IF FStep = CompleteState THEN
    FCompletedSequence := FCaptureStatus.SequenceId;
END_IF;
IF FStep >= LateChildProgress THEN
    FStatusRefreshMatches := (Snapshot.Execution.State = E_State.Completed)
        AND Snapshot.Execution.Completed AND NOT Snapshot.Execution.Ready
        AND (Snapshot.Execution.Result = FExpectedFinalResult)
        AND (Snapshot.TestCaseCountTotal = 2) AND (Snapshot.TestCaseCountRunning = 0);
    IF LateResetChildren THEN
        FStatusRefreshMatches := FStatusRefreshMatches AND Snapshot.Execution.Error
            AND (Snapshot.TestCaseCountCompleted = 1) AND (Snapshot.TestCaseCountError = 1)
            AND (Snapshot.TestCaseCountIdle = 1) AND (Snapshot.TestCaseCountPassed = 0);
    ELSE
        FStatusRefreshMatches := FStatusRefreshMatches AND NOT Snapshot.Execution.Error
            AND (Snapshot.TestCaseCountCompleted = 2) AND (Snapshot.TestCaseCountPassed = 2)
            AND (Snapshot.TestCaseCountIdle = 0) AND (Snapshot.TestCaseCountError = 0);
    END_IF;
    FPublicationMatches := FPublicationMatches AND (FCaptureStatus.SequenceId = FCompletedSequence);
END_IF;
IF (FStep = ReleaseReservations) OR (FStep = QuietAfterRelease)
    OR ((FStep = ResetOutcome) AND NOT LateResetChildren) THEN
    Released := FSubject.FreeReservedEvents();
    FCleanupMatches := Released
        AND (FSubject.ReservedEntryCount = 0) AND (FCapture.ReservedEntryCount = 0)
        AND (FSubject.State = ExpectedState) AND (FSubject.Result = ExpectedResult);
END_IF;

IF FExpectCompletion THEN
    FPublicationMatches := FPublicationMatches AND (FCaptureStatus.SequenceId = FCompletedSequence);
END_IF;
END_METHOD

END_FUNCTION_BLOCK

// ---- SelfTests/TestCases/TestSuite_TestSuiteLifecycle/Test_SuiteReservationRelease.TcPOU
{region 'Documentation'}
(*!
<summary>Verifies Suite release delegation, partial success, zero-own-budget cleanup and idempotent retry.</summary>
<description>

Boundary under test

The Suite uses the real local EventBuffer for its own contribution. Controlled children retain
local reservation markers only; they deliberately do not reproduce global reservation accounting.
The test checks that every child is called even if the first rejects release and that the Suite
still releases its own contribution. Global child-budget arithmetic belongs to capacity tests.

Retry and lifecycle

A failed child keeps its marker. A later successful retry releases it without re-releasing
already cleared contributions. Cleanup also visits children when the Suite's own count is zero.
None of these calls may issue child lifecycle requests, change owner state or restart execution.
</description>
*)
{endregion}
FUNCTION_BLOCK Test_SuiteReservationRelease EXTENDS TestCaseBase
VAR
    FSubjectParent : I_RunControl;
    FSubject : TestSuiteLifecycleProbe;
    FHelper : SuiteOrchestratorDouble;
    FCapture : EventBuffer;
    FEvents : ARRAY[1..CaptureLength] OF ST_Event;
    FCaptureFifo : ST_FifoStatus;
    FCaptureStatus : ST_EventBufferStatus;
    FChildView : ST_OrchestrationObservation;
    FStep : INT;
    FStepChecked : BOOL;
    FQuietSequence : UDINT;
    FDelegation : AssertTrue;
    FDelegationMatches : BOOL := TRUE;
    FOwnRelease : AssertTrue;
    FOwnReleaseMatches : BOOL := TRUE;
    FIdempotence : AssertTrue;
    FIdempotenceMatches : BOOL := TRUE;
    FNoLifecycleEffects : AssertTrue;
    FNoLifecycleEffectsMatches : BOOL := TRUE;
    FChildCalls : AssertTrue;
    FChildCallsMatches : BOOL := TRUE;
END_VAR
VAR CONSTANT
    CaptureLength : UINT := 64;
    ReservationMarker : UINT := 1;
    Setup : INT := 0;
    ResetRequested : INT := 1;
    FinishReset : INT := 2;
    ReserveAll : INT := 3;
    PartialRelease : INT := 4;
    RetryRelease : INT := 5;
    ReleaseWithZeroOwnCount : INT := 6;
    RepeatRelease : INT := 7;
    Done : INT := 8;
END_VAR

SUPER^();

{region 'Documentation'}
(*!
<summary>Contributes only the checking Assertions, not the intentionally controlled subject results.</summary>
*)
{endregion}
METHOD PROTECTED AggregateResults
VAR_INPUT
    Aggregator : I_ResultAggregator; //! Borrowed result sink owned by the outer Test Case; add this test's checking Assertions without resetting or retaining the sink.
END_VAR
Aggregator.AddProvider(Provider := FDelegation);
Aggregator.AddProvider(Provider := FOwnRelease);
Aggregator.AddProvider(Provider := FIdempotence);
Aggregator.AddProvider(Provider := FNoLifecycleEffects);
Aggregator.AddProvider(Provider := FChildCalls);
END_METHOD

{region 'Documentation'}
(*!
<summary>Supplies only the root identity; the root never executes this isolated subject.</summary>
*)
{endregion}
METHOD PUBLIC BindSubjectParent
VAR_INPUT
    Parent : I_RunControl; //! Borrowed identity parent retained for isolated subject initialization; keep the Run-Control alive through subject use.
END_VAR
FSubjectParent := Parent;
END_METHOD

{region 'Documentation'}
(*!
<summary>Initializes the checking Assertions; the scenario explicitly initializes its isolated subject.</summary>
*)
{endregion}
METHOD PROTECTED Configure
FPreparationStateCount := 0;
FTestStateCount := 1;
FDelegation.Initialize(Parent := THIS^,
    AssertionName := 'Delegation');
FOwnRelease.Initialize(Parent := THIS^,
    AssertionName := 'OwnRelease');
FIdempotence.Initialize(Parent := THIS^,
    AssertionName := 'Idempotence');
FNoLifecycleEffects.Initialize(Parent := THIS^,
    AssertionName := 'NoLifecycleEffects');
FChildCalls.Initialize(Parent := THIS^,
    AssertionName := 'ChildCalls');
END_METHOD

{region 'Documentation'}
(*!
<summary>No asynchronous test resource remains to stop.</summary>
*)
{endregion}
METHOD PROTECTED ProcessAbort
VAR_INPUT
    Enable : BOOL; //! Phase permission supplied by the owning Test Case; FALSE does not authorize progression, while observation may continue.
END_VAR
IF Enable THEN
    CompleteAbort();
END_IF;
END_METHOD

{region 'Documentation'}
(*!
<summary>Checks each cleanup checkpoint before advancing; failures remain latched.</summary>
*)
{endregion}
METHOD PROTECTED ProcessAssertions
VAR_INPUT
    Enable : BOOL; //! Phase permission supplied by the owning Test Case; FALSE does not authorize progression, while observation may continue.
END_VAR
FDelegation(Enable := Enable,
    State := State,
    IN := FDelegationMatches);
FOwnRelease(Enable := Enable,
    State := State,
    IN := FOwnReleaseMatches);
FIdempotence(Enable := Enable,
    State := State,
    IN := FIdempotenceMatches);
FNoLifecycleEffects(Enable := Enable,
    State := State,
    IN := FNoLifecycleEffectsMatches);
FChildCalls(Enable := Enable,
    State := State,
    IN := FChildCallsMatches);
IF Enable THEN
    FStepChecked := TRUE;
END_IF;
END_METHOD

{region 'Documentation'}
(*!
<summary>No resource Preparation is required for this controlled owner scenario.</summary>
*)
{endregion}
METHOD PROTECTED ProcessPreparations
VAR_INPUT
    // SA0033: Required override; the scenario has no Preparation phase.
    {attribute 'analysis' := '-33'}
    Enable : BOOL; //! Phase permission supplied by the owning Test Case; FALSE does not authorize progression, while observation may continue.
END_VAR
END_METHOD

{region 'Documentation'}
(*!
<summary>Restarts the test script and clears checking Assertions; subject setup belongs to the next test attempt.</summary>
*)
{endregion}
METHOD PROTECTED ProcessReset
FStep := Setup;
FStepChecked := FALSE;
FQuietSequence := 0;
FDelegationMatches := TRUE;
FOwnReleaseMatches := TRUE;
FIdempotenceMatches := TRUE;
FNoLifecycleEffectsMatches := TRUE;
FChildCallsMatches := TRUE;
FDelegation.Reset();
FOwnRelease.Reset();
FIdempotence.Reset();
FNoLifecycleEffects.Reset();
FChildCalls.Reset();
CompleteReset();
END_METHOD

{region 'Documentation'}
(*!
<summary>Advances the explicit test script with at most one subject FB call per active PLC cycle.</summary>
*)
{endregion}
METHOD PROTECTED ProcessTests
VAR_INPUT
    Enable : BOOL; //! Phase permission supplied by the owning Test Case; FALSE does not authorize progression, while observation may continue.
END_VAR
IF NOT Enable THEN
    RETURN;
END_IF;
IF FStepChecked THEN
    FStep := FStep + 1;
    FStepChecked := FALSE;
END_IF;
IF FStep = Done THEN
    CompleteTests();
    RETURN;
END_IF;
RunStep();
END_METHOD

{region 'Documentation'}
(*!
<summary>Exercises a bounded cleanup sequence in Idle, recording each concrete child release attempt.</summary>
*)
{endregion}
METHOD PRIVATE RunStep
VAR
    Config : ST_TestSuiteConfig;
    FirstChild : I_TestCase;
    SecondChild : I_TestCase;
    FirstCalls : ST_OrchestrationCalls;
    SecondCalls : ST_OrchestrationCalls;
    ExpectedState : E_State;
    ExpectedTask : E_OrchestratorTask;
    Released : BOOL;
END_VAR
IF FStep = Setup THEN
    IF NOT FCapture.Initialize(Buffer := FEvents,
        FifoControl := FCaptureFifo,
        Status := FCaptureStatus) THEN
        Error(Message := 'Suite release capture could not be initialized.');
        RETURN;
    END_IF;
    FHelper.BeginScenario();
    FSubject.Bind(Publisher := FCapture,
        Helper := FHelper);
    IF NOT FSubject.Initialize(Parent := FSubjectParent,
        SuiteName := 'ReleaseSubject',
        Config := Config) THEN
        Error(Message := 'Suite release subject could not be initialized.');
        RETURN;
    END_IF;
END_IF;
FirstChild := FSubject.GetTestCase(Index := FSubject.ChildArrayLowerBound);
SecondChild := FSubject.GetTestCase(Index := FSubject.ChildArrayLowerBound + 1);
ExpectedState := E_State.Idle;
ExpectedTask := E_OrchestratorTask.Idle;

CASE FStep OF
    Setup:
        FChildView.State := E_State.Uninitialized;
        FChildView.Result := E_Result.NotEvaluated;
        FChildView.Ready := FALSE;
        FChildView.Complete := FALSE;
        ExpectedState := E_State.Uninitialized;

    ResetRequested:
        IF FSubject.ReserveResetEvents() <> E_EventReservationResult.Accepted THEN
            Error(Message := 'Suite release fixture Reset reservation was rejected.');
            RETURN;
        END_IF;
        FSubject.RequestReset();
        FChildView.State := E_State.Reset;
        ExpectedState := E_State.Reset;
        ExpectedTask := E_OrchestratorTask.Reset;

    FinishReset:
        FHelper.SetObservation(Ready := TRUE,
            ResetFinished := TRUE);
        FChildView.State := E_State.Idle;
        FChildView.Ready := TRUE;

    ReserveAll:
        IF FSubject.ReserveExecutionEvents() <> E_EventReservationResult.Accepted THEN
            Error(Message := 'Suite release fixture execution reservation was rejected.');
            RETURN;
        END_IF;
        IF FirstChild.ReserveExecutionEvents() <> E_EventReservationResult.Accepted THEN
            Error(Message := 'First controlled child reservation was rejected.');
            RETURN;
        END_IF;
        IF SecondChild.ReserveExecutionEvents() <> E_EventReservationResult.Accepted THEN
            Error(Message := 'Second controlled child reservation was rejected.');
            RETURN;
        END_IF;
        FOwnReleaseMatches := (FSubject.ReservedEntryCount > 0)
            AND (FCapture.ReservedEntryCount = FSubject.ReservedEntryCount);
        FDelegationMatches := (FirstChild.ReservedEntryCount = ReservationMarker)
            AND (SecondChild.ReservedEntryCount = ReservationMarker);

    PartialRelease:
        FSubject.SetChildReleaseResponses(FirstSucceeds := FALSE);
        Released := FSubject.FreeReservedEvents();
        FirstCalls := FSubject.GetChildCalls(Index := FSubject.ChildArrayLowerBound);
        SecondCalls := FSubject.GetChildCalls(Index := FSubject.ChildArrayLowerBound + 1);
        FDelegationMatches := NOT Released AND (FirstCalls.FreeCount = 1) AND (SecondCalls.FreeCount = 1)
            AND (FirstChild.ReservedEntryCount = ReservationMarker) AND (SecondChild.ReservedEntryCount = 0)
            AND (FirstCalls.ReleasedEntryCount = 0) AND (SecondCalls.ReleasedEntryCount = ReservationMarker);
        FOwnReleaseMatches := (FSubject.ReservedEntryCount = 0) AND (FCapture.ReservedEntryCount = 0);

    RetryRelease:
        FSubject.SetChildReleaseResponses();
        Released := FSubject.FreeReservedEvents();
        FirstCalls := FSubject.GetChildCalls(Index := FSubject.ChildArrayLowerBound);
        SecondCalls := FSubject.GetChildCalls(Index := FSubject.ChildArrayLowerBound + 1);
        FDelegationMatches := Released AND (FirstCalls.FreeCount = 2) AND (SecondCalls.FreeCount = 2)
            AND (FirstChild.ReservedEntryCount = 0) AND (SecondChild.ReservedEntryCount = 0);
        FIdempotenceMatches := (FirstCalls.ReleasedEntryCount = ReservationMarker)
            AND (SecondCalls.ReleasedEntryCount = ReservationMarker);

    ReleaseWithZeroOwnCount:
        IF FirstChild.ReserveResetEvents() <> E_EventReservationResult.Accepted THEN
            Error(Message := 'First controlled child Reset reservation was rejected.');
            RETURN;
        END_IF;
        IF SecondChild.ReserveResetEvents() <> E_EventReservationResult.Accepted THEN
            Error(Message := 'Second controlled child Reset reservation was rejected.');
            RETURN;
        END_IF;
        FOwnReleaseMatches := FSubject.ReservedEntryCount = 0;
        Released := FSubject.FreeReservedEvents();
        FirstCalls := FSubject.GetChildCalls(Index := FSubject.ChildArrayLowerBound);
        SecondCalls := FSubject.GetChildCalls(Index := FSubject.ChildArrayLowerBound + 1);
        FDelegationMatches := Released AND (FirstCalls.FreeCount = 3) AND (SecondCalls.FreeCount = 3)
            AND (FirstChild.ReservedEntryCount = 0) AND (SecondChild.ReservedEntryCount = 0);
        FIdempotenceMatches := (FirstCalls.ReleasedEntryCount = 2 * ReservationMarker)
            AND (SecondCalls.ReleasedEntryCount = 2 * ReservationMarker);

    RepeatRelease:
        Released := FSubject.FreeReservedEvents();
        FirstCalls := FSubject.GetChildCalls(Index := FSubject.ChildArrayLowerBound);
        SecondCalls := FSubject.GetChildCalls(Index := FSubject.ChildArrayLowerBound + 1);
        FDelegationMatches := Released AND (FirstCalls.FreeCount = 4) AND (SecondCalls.FreeCount = 4);
        FIdempotenceMatches := (FirstCalls.ReleasedEntryCount = 2 * ReservationMarker)
            AND (SecondCalls.ReleasedEntryCount = 2 * ReservationMarker)
            AND (FirstChild.ReservedEntryCount = 0) AND (SecondChild.ReservedEntryCount = 0)
            AND (FSubject.ReservedEntryCount = 0) AND (FCapture.ReservedEntryCount = 0);
ELSE
    Error(Message := 'Unexpected Suite release test step.');
    RETURN;
END_CASE;

FSubject.SetChildObservation(Observation := FChildView);
FSubject();
FirstCalls := FSubject.GetChildCalls(Index := FSubject.ChildArrayLowerBound);
SecondCalls := FSubject.GetChildCalls(Index := FSubject.ChildArrayLowerBound + 1);
FNoLifecycleEffectsMatches := (FSubject.State = ExpectedState)
    AND (FSubject.Result = E_Result.NotEvaluated) AND (FHelper.CurrentTask = ExpectedTask)
    AND (FirstChild.State = FChildView.State) AND (SecondChild.State = FChildView.State)
    AND (FirstCalls.StartCount = 0) AND (FirstCalls.ResetCount = 0) AND (FirstCalls.AbortCount = 0)
    AND (SecondCalls.StartCount = 0) AND (SecondCalls.ResetCount = 0) AND (SecondCalls.AbortCount = 0);
FChildCallsMatches := FSubject.ChildBodyCallsMatch
    AND (FSubject.ChildCallCount = INT_TO_UINT(FStep + 1))
    AND (FHelper.ExecuteCount = INT_TO_UINT(FStep + 1));
IF FStep = FinishReset THEN
    FQuietSequence := FCaptureStatus.SequenceId;
END_IF;
IF FStep >= ReserveAll THEN
    FNoLifecycleEffectsMatches := FNoLifecycleEffectsMatches AND FSubject.IsReady
        AND (FCaptureStatus.SequenceId = FQuietSequence) AND (FCaptureStatus.LostEventCount = 0);
END_IF;
END_METHOD

END_FUNCTION_BLOCK

// ---- SelfTests/TestCases/TestSuite_TestSuiteLifecycle/Test_SuiteRealComposition.TcPOU
{region 'Documentation'}
(*!
<summary>Runs one real Suite composition twice with a lifecycle Reset between executions.</summary>
<description>

Real boundaries

The subject owns two minimal real Test Cases and the production Orchestrator.
The outer test supplies only parent Reset/Start requests and the Suite's own event budget.
It does not manufacture child or helper observations.

Repeat and isolation

Initialize runs once. Both executions must finish Passed; Reset must restore Idle,
NotEvaluated and readiness without rebuilding the collection. While Reset remains active,
the parent repeats RequestReset on each waiting call; real child/helper progress must survive.
All subject producers share a local capture retained across both runs.
Each child's finalization must precede the Suite's finalization, and parent release
must leave no held reservations. Detailed scheduling remains in its dedicated tests.
</description>
*)
{endregion}
FUNCTION_BLOCK Test_SuiteRealComposition EXTENDS TestCaseBase
VAR
    FSubjectParent : I_RunControl;
    FSubject : SuiteIntegrationSubject;
    FCapture : EventBuffer;
    FEvents : ARRAY[1..CaptureLength] OF ST_Event;
    FCaptureFifo : ST_FifoStatus;
    FCaptureStatus : ST_EventBufferStatus;
    FStep : INT;
    FCompletedRuns : UINT;
    FFinalChecksEvaluated : BOOL;
    FReadiness : AssertTrue;
    FReadinessMatches : BOOL := TRUE;
    FCompletion : AssertTrue;
    FCompletionMatches : BOOL := TRUE;
    FRepeat : AssertTrue;
    FRepeatMatches : BOOL := TRUE;
    FReservations : AssertTrue;
    FReservationsMatches : BOOL := TRUE;
    FChildCalls : AssertTrue;
    FChildCallsMatches : BOOL := TRUE;
    FEventStream : AssertTrue;
    FEventStreamMatches : BOOL := TRUE;
END_VAR
VAR CONSTANT
    CaptureLength : UINT := 256;
    ExpectedChildCount : UINT := 2;
    RequiredRuns : UINT := 2;
    Setup : INT := 0;
    ResetRequested : INT := 1;
    WaitForReadiness : INT := 2;
    StartRequested : INT := 3;
    WaitForCompletion : INT := 4;
    Finish : INT := 5;
END_VAR

SUPER^();

{region 'Documentation'}
(*!
<summary>Contributes only the checking Assertions, not the intentionally controlled subject results.</summary>
*)
{endregion}
METHOD PROTECTED AggregateResults
VAR_INPUT
    Aggregator : I_ResultAggregator; //! Borrowed result sink owned by the outer Test Case; add this test's checking Assertions without resetting or retaining the sink.
END_VAR
Aggregator.AddProvider(Provider := FReadiness);
Aggregator.AddProvider(Provider := FCompletion);
Aggregator.AddProvider(Provider := FRepeat);
Aggregator.AddProvider(Provider := FReservations);
Aggregator.AddProvider(Provider := FChildCalls);
Aggregator.AddProvider(Provider := FEventStream);
END_METHOD

{region 'Documentation'}
(*!
<summary>Supplies only the root identity; the root never executes this isolated subject.</summary>
*)
{endregion}
METHOD PUBLIC BindSubjectParent
VAR_INPUT
    Parent : I_RunControl; //! Borrowed identity parent retained for isolated subject initialization; keep the Run-Control alive through subject use.
END_VAR
FSubjectParent := Parent;
END_METHOD

{region 'Documentation'}
(*!
<summary>Checks exact finalization counts and latest child-before-owner event order across both executions.</summary>
*)
{endregion}
METHOD PRIVATE CheckEventStream
VAR
    Index : UINT;
    SuiteResults : UINT;
    SuiteAggregations : UINT;
    SuiteCompletions : UINT;
    FirstResults : UINT;
    SecondResults : UINT;
    FirstCompletions : UINT;
    SecondCompletions : UINT;
    SuiteResultSequence : UDINT;
    SuiteAggregationSequence : UDINT;
    SuiteCompletionSequence : UDINT;
    FirstCompletionSequence : UDINT;
    SecondCompletionSequence : UDINT;
    FirstChild : I_TestCase;
    SecondChild : I_TestCase;
END_VAR
FirstChild := FSubject.GetTestCase(Index := FSubject.ChildArrayLowerBound);
SecondChild := FSubject.GetTestCase(Index := FSubject.ChildArrayLowerBound + 1);
FOR Index := 1 TO CaptureLength DO
    IF FEvents[Index].SequenceId = 0 THEN
        CONTINUE;
    END_IF;
    FEventStreamMatches := FEventStreamMatches
        AND (FEvents[Index].Severity <> E_EventSeverity.Error);
    IF FEvents[Index].Name = FSubject.Name THEN
        CASE FEvents[Index].EventType OF
            E_EventType.Result:
                SuiteResults := SuiteResults + 1;
                SuiteResultSequence := FEvents[Index].SequenceId;
                FEventStreamMatches := FEventStreamMatches AND (FEvents[Index].Result = E_Result.Passed);
            E_EventType.Aggregation:
                SuiteAggregations := SuiteAggregations + 1;
                SuiteAggregationSequence := FEvents[Index].SequenceId;
            E_EventType.StateTransition:
                IF FEvents[Index].State = E_State.Completed THEN
                    SuiteCompletions := SuiteCompletions + 1;
                    SuiteCompletionSequence := FEvents[Index].SequenceId;
                END_IF;
        END_CASE;
    ELSIF FEvents[Index].Name = FirstChild.Name THEN
        IF FEvents[Index].EventType = E_EventType.Result THEN
            FirstResults := FirstResults + 1;
        ELSIF (FEvents[Index].EventType = E_EventType.StateTransition)
            AND (FEvents[Index].State = E_State.Completed) THEN
            FirstCompletions := FirstCompletions + 1;
            FirstCompletionSequence := FEvents[Index].SequenceId;
        END_IF;
    ELSIF FEvents[Index].Name = SecondChild.Name THEN
        IF FEvents[Index].EventType = E_EventType.Result THEN
            SecondResults := SecondResults + 1;
        ELSIF (FEvents[Index].EventType = E_EventType.StateTransition)
            AND (FEvents[Index].State = E_State.Completed) THEN
            SecondCompletions := SecondCompletions + 1;
            SecondCompletionSequence := FEvents[Index].SequenceId;
        END_IF;
    END_IF;
END_FOR;
FEventStreamMatches := FEventStreamMatches
    AND (SuiteResults = FCompletedRuns) AND (SuiteAggregations = FCompletedRuns)
    AND (SuiteCompletions = FCompletedRuns)
    AND (FirstResults = FCompletedRuns) AND (SecondResults = FCompletedRuns)
    AND (FirstCompletions = FCompletedRuns) AND (SecondCompletions = FCompletedRuns)
    AND (FirstCompletionSequence < SuiteResultSequence)
    AND (SecondCompletionSequence < SuiteResultSequence)
    AND (SuiteResultSequence < SuiteAggregationSequence)
    AND (SuiteAggregationSequence < SuiteCompletionSequence);
END_METHOD

{region 'Documentation'}
(*!
<summary>Initializes the checking Assertions; the scenario explicitly initializes its isolated subject.</summary>
*)
{endregion}
METHOD PROTECTED Configure
FPreparationStateCount := 0;
FTestStateCount := 1;
FReadiness.Initialize(Parent := THIS^,
    AssertionName := 'Readiness');
FCompletion.Initialize(Parent := THIS^,
    AssertionName := 'Completion');
FRepeat.Initialize(Parent := THIS^,
    AssertionName := 'Repeat');
FReservations.Initialize(Parent := THIS^,
    AssertionName := 'Reservations');
FChildCalls.Initialize(Parent := THIS^,
    AssertionName := 'ChildCalls');
FEventStream.Initialize(Parent := THIS^,
    AssertionName := 'EventStream');
END_METHOD

{region 'Documentation'}
(*!
<summary>No asynchronous test resource remains to stop.</summary>
*)
{endregion}
METHOD PROTECTED ProcessAbort
VAR_INPUT
    Enable : BOOL; //! Phase permission supplied by the owning Test Case; FALSE does not authorize progression, while observation may continue.
END_VAR
IF Enable THEN
    CompleteAbort();
END_IF;
END_METHOD

{region 'Documentation'}
(*!
<summary>Keeps every observation across both runs; final checks must evaluate before ending the outer Test Case.</summary>
*)
{endregion}
METHOD PROTECTED ProcessAssertions
VAR_INPUT
    Enable : BOOL; //! Phase permission supplied by the owning Test Case; FALSE does not authorize progression, while observation may continue.
END_VAR
FReadiness(Enable := Enable,
    State := State,
    IN := FReadinessMatches);
FCompletion(Enable := Enable,
    State := State,
    IN := FCompletionMatches);
FRepeat(Enable := Enable,
    State := State,
    IN := FRepeatMatches);
FReservations(Enable := Enable,
    State := State,
    IN := FReservationsMatches);
FChildCalls(Enable := Enable,
    State := State,
    IN := FChildCallsMatches);
FEventStream(Enable := Enable,
    State := State,
    IN := FEventStreamMatches);
IF Enable AND (FStep = Finish) THEN
    FFinalChecksEvaluated := TRUE;
END_IF;
END_METHOD

{region 'Documentation'}
(*!
<summary>No resource Preparation is required for this controlled owner scenario.</summary>
*)
{endregion}
METHOD PROTECTED ProcessPreparations
VAR_INPUT
    // SA0033: Required override; the scenario has no Preparation phase.
    {attribute 'analysis' := '-33'}
    Enable : BOOL; //! Phase permission supplied by the owning Test Case; FALSE does not authorize progression, while observation may continue.
END_VAR
END_METHOD

{region 'Documentation'}
(*!
<summary>Restarts the test script and clears checking Assertions; subject setup belongs to the next test attempt.</summary>
*)
{endregion}
METHOD PROTECTED ProcessReset
FStep := Setup;
FCompletedRuns := 0;
FFinalChecksEvaluated := FALSE;
FReadinessMatches := TRUE;
FCompletionMatches := TRUE;
FRepeatMatches := TRUE;
FReservationsMatches := TRUE;
FChildCallsMatches := TRUE;
FEventStreamMatches := TRUE;
FReadiness.Reset();
FCompletion.Reset();
FRepeat.Reset();
FReservations.Reset();
FChildCalls.Reset();
FEventStream.Reset();
CompleteReset();
END_METHOD

{region 'Documentation'}
(*!
<summary>Advances the explicit test script with at most one subject FB call per active PLC cycle.</summary>
*)
{endregion}
METHOD PROTECTED ProcessTests
VAR_INPUT
    Enable : BOOL; //! Phase permission supplied by the owning Test Case; FALSE does not authorize progression, while observation may continue.
END_VAR
IF NOT Enable THEN
    RETURN;
END_IF;
IF (FStep = Finish) AND FFinalChecksEvaluated THEN
    CompleteTests();
    RETURN;
END_IF;
RunStep();
END_METHOD

{region 'Documentation'}
(*!
<summary>Performs the parent-owned release and checks global and per-child accounting, including repeated release.</summary>
*)
{endregion}
METHOD PRIVATE ReleaseAndCheck
VAR
    FirstChild : I_TestCase;
    SecondChild : I_TestCase;
    Released : BOOL;
END_VAR
Released := FSubject.FreeReservedEvents();
FReservationsMatches := FReservationsMatches AND Released;
Released := FSubject.FreeReservedEvents();
FirstChild := FSubject.GetTestCase(Index := FSubject.ChildArrayLowerBound);
SecondChild := FSubject.GetTestCase(Index := FSubject.ChildArrayLowerBound + 1);
FReservationsMatches := FReservationsMatches AND Released
    AND (FSubject.ReservedEntryCount = 0)
    AND (FirstChild.ReservedEntryCount = 0) AND (SecondChild.ReservedEntryCount = 0)
    AND (FCapture.ReservedEntryCount = 0);
END_METHOD

{region 'Documentation'}
(*!
<summary>Issues parent requests once and otherwise lets the real composition progress one FB call per PLC cycle.</summary>
*)
{endregion}
METHOD PRIVATE RunStep
VAR
    Config : ST_TestSuiteConfig;
    Snapshot : ST_TestSuiteStatus;
    FirstChild : I_TestCase;
    SecondChild : I_TestCase;
END_VAR
CASE FStep OF
    Setup:
        IF NOT FCapture.Initialize(Buffer := FEvents,
            FifoControl := FCaptureFifo,
            Status := FCaptureStatus) THEN
            Error(Message := 'Real Suite composition capture initialization failed.');
            RETURN;
        END_IF;
        FSubject.BindPublisher(Publisher := FCapture);
        IF NOT FSubject.Initialize(Parent := FSubjectParent,
            SuiteName := 'RealComposition',
            Config := Config) THEN
            Error(Message := 'Real Suite composition initialization failed.');
            RETURN;
        END_IF;
        FStep := ResetRequested;

    ResetRequested:
        IF FSubject.ReserveResetEvents() <> E_EventReservationResult.Accepted THEN
            Error(Message := 'Real Suite composition Reset reservation was rejected.');
            RETURN;
        END_IF;
        FSubject.RequestReset();
        FStep := WaitForReadiness;

    StartRequested:
        IF FSubject.ReserveExecutionEvents() <> E_EventReservationResult.Accepted THEN
            Error(Message := 'Real Suite composition execution reservation was rejected.');
            RETURN;
        END_IF;
        FSubject.RequestStart();
        FStep := WaitForCompletion;

    WaitForReadiness:
        IF FSubject.IsResetting THEN
            FSubject.RequestReset();
        END_IF;

    WaitForCompletion, Finish:
        // Waiting retains real child/helper timing; the outer Test Case timeout bounds a stalled subject.
ELSE
    Error(Message := 'Unexpected real Suite composition test step.');
    RETURN;
END_CASE;

FSubject();
FChildCallsMatches := FChildCallsMatches AND FSubject.ChildCallsMatch;
FRepeatMatches := FRepeatMatches AND (FSubject.ConfigureCount = 1)
    AND (FSubject.ChildCount = ExpectedChildCount);
FEventStreamMatches := FEventStreamMatches AND (FCaptureStatus.LostEventCount = 0);
Snapshot := FSubject.Status;

CASE FStep OF
    WaitForReadiness:
        IF FSubject.HasError THEN
            Error(Message := 'Real Suite composition failed during Reset.');
            RETURN;
        END_IF;
        IF FSubject.IsReady THEN
            FReadinessMatches := FReadinessMatches AND FSubject.IsIdle
                AND (FSubject.Result = E_Result.NotEvaluated)
                AND (Snapshot.TestCaseCountIdle = ExpectedChildCount)
                AND (Snapshot.TestCaseCountCompleted = 0);
            ReleaseAndCheck();
            FStep := StartRequested;
        END_IF;

    WaitForCompletion:
        IF FSubject.IsComplete THEN
            FirstChild := FSubject.GetTestCase(Index := FSubject.ChildArrayLowerBound);
            SecondChild := FSubject.GetTestCase(Index := FSubject.ChildArrayLowerBound + 1);
            FCompletionMatches := FCompletionMatches
                AND (FSubject.Result = E_Result.Passed)
                AND (Snapshot.TestCaseCountCompleted = ExpectedChildCount)
                AND (Snapshot.TestCaseCountPassed = ExpectedChildCount)
                AND (Snapshot.TestCaseCountFailed = 0) AND (Snapshot.TestCaseCountError = 0)
                AND FirstChild.IsComplete AND SecondChild.IsComplete
                AND (FirstChild.Result = E_Result.Passed) AND (SecondChild.Result = E_Result.Passed);
            FCompletedRuns := FCompletedRuns + 1;
            ReleaseAndCheck();
            CheckEventStream();
            IF FCompletedRuns = RequiredRuns THEN
                FStep := Finish;
            ELSE
                FStep := ResetRequested;
            END_IF;
        END_IF;
END_CASE;
END_METHOD

END_FUNCTION_BLOCK

// ---- SelfTests/TestCases/TestSuite_TestSuiteLifecycle/Helper/SuiteIntegrationSubject.TcPOU
{region 'Documentation'}
(*!
<summary>Composes two minimal real Test Cases with the real production Orchestrator.</summary>
<description>
Only publisher binding and call counters are added for observation.
The inherited base and real helper own all transitions, requests and reservations.
Children are initialized once in Configure, then Reset and executed twice without rebinding.
</description>
*)
{endregion}
FUNCTION_BLOCK SuiteIntegrationSubject EXTENDS TestSuiteBase
VAR
    FFirst : SuiteIntegrationChild;
    FSecond : SuiteIntegrationChild;
    FTestCases : ARRAY[4..6] OF I_TestCase;
    FRealOrchestrator : OrchestratorProbe;
    FBodyCallCount : UDINT;
    FConfigureCount : UINT;
END_VAR

FBodyCallCount := FBodyCallCount + 1;
SUPER^();

{region 'Documentation'}
(*!
<summary>Binds every producer before Initialize; never modifies the global publisher.</summary>
*)
{endregion}
METHOD PUBLIC BindPublisher
VAR_INPUT
    Publisher : I_EventPublisher; //! Nonzero isolated event publisher retained before subject initialization; keep it alive through all subject use.
END_VAR
FEventPublisher := Publisher;
FRealOrchestrator.BindPublisher(Publisher := Publisher);
FOrchestrator := FRealOrchestrator;
FFirst.BindPublisher(Publisher := Publisher);
FSecond.BindPublisher(Publisher := Publisher);
FBodyCallCount := 0;
FConfigureCount := 0;
END_METHOD

{region 'Documentation'}
(*!
<summary>Confirms one concrete child call per Suite call, including Reset and Completed.</summary>
*)
{endregion}
{attribute 'monitoring' := 'call'}
PROPERTY PUBLIC ChildCallsMatch : BOOL //! Confirms one concrete child call per Suite call, including Reset and Completed.
GET
ChildCallsMatch := (FFirst.BodyCallCount = FBodyCallCount) AND (FSecond.BodyCallCount = FBodyCallCount);
END_GET
END_PROPERTY

{region 'Documentation'}
(*!
<summary>Initializes and registers two real children serially in a shifted array with one unused slot.</summary>
*)
{endregion}
METHOD PROTECTED Configure
VAR_IN_OUT
    // SA0167: Borrowed setup builder; no temporary instance is created.
    {attribute 'analysis' := '-167'}
    Builder : TestSuiteConfigurationBuilder; //! Borrowed owner configuration builder used only during this Configure call; register this owner's concrete children.
END_VAR
VAR
    Config : ST_TestCaseConfig;
END_VAR
FConfigureCount := FConfigureCount + 1;
Builder.Initialize(Mode := E_OrchestrationMode.Serial,
    TestCases := FTestCases);
FFirst.Initialize(Parent := THIS^,
    TestName := 'First',
    Config := Config);
FSecond.Initialize(Parent := THIS^,
    TestName := 'Second',
    Config := Config);
Builder.Register(TestCase := FFirst);
Builder.Register(TestCase := FSecond);
END_METHOD

{region 'Documentation'}
(*!
<summary>Distinguishes Reset/repeat from reinitializing the subject.</summary>
*)
{endregion}
{attribute 'monitoring' := 'call'}
PROPERTY PUBLIC ConfigureCount : UINT //! Distinguishes Reset/repeat from reinitializing the subject.
GET
ConfigureCount := FConfigureCount;
END_GET
END_PROPERTY

{region 'Documentation'}
(*!
<summary>Resolves the actual registered array index without executing the child.</summary>
*)
{endregion}
METHOD PUBLIC GetTestCase : I_TestCase //! Typed child interface at the original array index; zero when no entry is available.
VAR_INPUT
    Index : DINT; //! Original occupied child-array index, rather than an ordinal position.
END_VAR
GetTestCase := 0;
IF (ChildCount = 0) OR (Index < ChildArrayLowerBound)
    OR (DINT_TO_LINT(Index) >= DINT_TO_LINT(ChildArrayLowerBound) + UINT_TO_LINT(ChildCount)) THEN
    RETURN;
END_IF;
GetTestCase := FTestCases[Index];
END_METHOD

{region 'Documentation'}
(*!
<summary>Calls both children once per initialized Suite call; the helper requests their lifecycle actions.</summary>
*)
{endregion}
METHOD PROTECTED ProcessTestCases
FFirst();
FSecond();
END_METHOD

END_FUNCTION_BLOCK

// ---- SelfTests/TestCases/TestSuite_TestSuiteLifecycle/Helper/SuiteIntegrationChild.TcPOU
{region 'Documentation'}
(*!
<summary>Exercises the successful framework lifecycle with one Boolean Assertion.</summary>
*)
{endregion}
FUNCTION_BLOCK SuiteIntegrationChild EXTENDS TestCaseBase
VAR
    FSuccess : AssertTrue;
    FBodyCallCount : UDINT;
    FActual : BOOL;
    FCheckPerformed : BOOL;
END_VAR

FBodyCallCount := FBodyCallCount + 1;
SUPER^();

{region 'Documentation'}
(*!
<summary>Contributes the one Assertion without executing or resetting it.</summary>
*)
{endregion}
METHOD PROTECTED AggregateResults
VAR_INPUT
    Aggregator : I_ResultAggregator; //! Borrowed result sink owned by the outer Test Case; add this test's checking Assertions without resetting or retaining the sink.
END_VAR
Aggregator.AddProvider(Provider := FSuccess);
END_METHOD

{region 'Documentation'}
(*!
<summary>Binds this real Test Case and its Assertion to the isolated capture before initialization.</summary>
*)
{endregion}
METHOD PUBLIC BindPublisher
VAR_INPUT
    Publisher : I_EventPublisher; //! Nonzero isolated event publisher retained before subject initialization; keep it alive through all subject use.
END_VAR
FEventPublisher := Publisher;
FSuccess.BindPublisher(Publisher := Publisher);
FBodyCallCount := 0;
END_METHOD

{region 'Documentation'}
(*!
<summary>Counts concrete FB calls since binding, including disabled lifecycle phases.</summary>
*)
{endregion}
{attribute 'monitoring' := 'call'}
PROPERTY PUBLIC BodyCallCount : UDINT //! Counts concrete FB calls since binding, including disabled lifecycle phases.
GET
BodyCallCount := FBodyCallCount;
END_GET
END_PROPERTY

{region 'Documentation'}
(*!
<summary>Includes the owned Assertion in the base initialization checks.</summary>
*)
{endregion}
METHOD PROTECTED CheckInitialization : BOOL //! TRUE when the inherited initialization check and this concrete fixture check both accept the setup.
CheckInitialization := FALSE;
IF NOT SUPER^.CheckInitialization() THEN
    RETURN;
END_IF;
IF NOT FSuccess.IsInitialized THEN
    RETURN;
END_IF;

CheckInitialization := TRUE;
END_METHOD

{region 'Documentation'}
(*!
<summary>Initializes the minimal integration scenario and its single Assertion.</summary>
*)
{endregion}
METHOD PROTECTED Configure
FPreparationStateCount := 0;
FTestStateCount := 1;
FActual := FALSE;
FCheckPerformed := FALSE;

FSuccess.Initialize(Parent := THIS^,
    AssertionName := 'Success');
END_METHOD

{region 'Documentation'}
(*!
<summary>Completes enabled aborts; the minimal integration scenario owns no resource actions.</summary>
*)
{endregion}
METHOD PROTECTED ProcessAbort
VAR_INPUT
    Enable : BOOL; //! Phase permission supplied by the owning Test Case; FALSE does not authorize progression, while observation may continue.
END_VAR
IF Enable THEN
    CompleteAbort();
END_IF;
END_METHOD

{region 'Documentation'}
(*!
<summary>Calls the Assertion even while disabled and records an actual evaluation.</summary>
*)
{endregion}
METHOD PROTECTED ProcessAssertions
VAR_INPUT
    Enable : BOOL; //! Phase permission supplied by the owning Test Case; FALSE does not authorize progression, while observation may continue.
END_VAR
FSuccess(Enable := Enable,
    State := State,
    IN := FActual);

IF Enable AND FSuccess.EvaluationActive THEN
    FCheckPerformed := TRUE;
END_IF;
END_METHOD

{region 'Documentation'}
(*!
<summary>No Preparation stage is configured for this minimal integration scenario.</summary>
*)
{endregion}
METHOD PROTECTED ProcessPreparations
VAR_INPUT
    // SA0033: Required override signature; this scenario has no preparation work.
    {attribute 'analysis' := '-33'}
    Enable : BOOL; //! Phase permission supplied by the owning Test Case; FALSE does not authorize progression, while observation may continue.
END_VAR
END_METHOD

{region 'Documentation'}
(*!
<summary>Clears scenario progress and requests Assertion reset before returning to Idle.</summary>
*)
{endregion}
METHOD PROTECTED ProcessReset
FActual := FALSE;
FCheckPerformed := FALSE;
FSuccess.Reset();
CompleteReset();
END_METHOD

{region 'Documentation'}
(*!
<summary>Supplies the success value, then completes on the call after evaluation.</summary>
*)
{endregion}
METHOD PROTECTED ProcessTests
VAR_INPUT
    Enable : BOOL; //! Phase permission supplied by the owning Test Case; FALSE does not authorize progression, while observation may continue.
END_VAR
IF NOT Enable THEN
    RETURN;
END_IF;

IF FCheckPerformed THEN
    CompleteTests();
ELSE
    FActual := TRUE;
END_IF;
END_METHOD

END_FUNCTION_BLOCK

// ---- SelfTests/TestCases/TestSuite_TestSuiteLifecycle/Test_SuiteMockRepeatedReset.TcPOU
{region 'Documentation'}
(*!
<summary>Verifies automatic mock Reset completion despite a second Reset request.</summary>
<description>
Each Reset retains its initial entry call, then reaches Idle on the next call even with
another request. A no-request call holds Idle before a second interval repeats the check.
The inherited mock owns all processing. A thin adapter only routes its events to local capture.
Checks cover coherent state/result/readiness, zero child counters, two Reset/Idle transitions,
reservation release and no lost events. Outer Assertions use the normal selftest publisher.
</description>
*)
{endregion}
FUNCTION_BLOCK Test_SuiteMockRepeatedReset EXTENDS TestCaseBase
VAR
    FSubjectParent : I_RunControl;
    FSubject : TestSuiteMockProbe;
    FCapture : EventBuffer;
    FEvents : ARRAY[1..CaptureLength] OF ST_Event;
    FCaptureFifo : ST_FifoStatus;
    FCaptureStatus : ST_EventBufferStatus;
    FStep : INT;
    FStepChecked : BOOL;
    FProgress : AssertTrue;
    FProgressMatches : BOOL := TRUE;
    FEvidence : AssertTrue;
    FEvidenceMatches : BOOL := TRUE;
END_VAR
VAR CONSTANT
    CaptureLength : UINT := 32;
    Setup : INT := 0;
    RequestFirst : INT := 1;
    RepeatFirst : INT := 2;
    HoldIdle : INT := 3;
    RequestAgain : INT := 4;
    RepeatAgain : INT := 5;
END_VAR

SUPER^();

{region 'Documentation'}
(*!
<summary>Contributes the checking Assertions and excludes the isolated subject.</summary>
*)
{endregion}
METHOD PROTECTED AggregateResults
VAR_INPUT
    Aggregator : I_ResultAggregator; //! Borrowed result sink; contribute checks without resetting or retaining it.
END_VAR
Aggregator.AddProvider(Provider := FProgress);
Aggregator.AddProvider(Provider := FEvidence);
END_METHOD

{region 'Documentation'}
(*!
<summary>Retains the root identity for the isolated mock subject.</summary>
*)
{endregion}
METHOD PUBLIC BindSubjectParent
VAR_INPUT
    Parent : I_RunControl; //! Borrowed root identity; keep alive throughout subject use.
END_VAR
FSubjectParent := Parent;
END_METHOD

{region 'Documentation'}
(*!
<summary>Initializes checks; subject initialization belongs to the active test scenario.</summary>
*)
{endregion}
METHOD PROTECTED Configure
FPreparationStateCount := 0;
FTestStateCount := 1;
FProgress.Initialize(Parent := THIS^,
    AssertionName := 'Progress');
FEvidence.Initialize(Parent := THIS^,
    AssertionName := 'Evidence');
END_METHOD

{region 'Documentation'}
(*!
<summary>Completes Abort immediately; no asynchronous resource is owned.</summary>
*)
{endregion}
METHOD PROTECTED ProcessAbort
VAR_INPUT
    Enable : BOOL; //! Authorizes completion of the active Abort phase.
END_VAR
IF Enable THEN
    CompleteAbort();
END_IF;
END_METHOD

{region 'Documentation'}
(*!
<summary>Checks the subject cycle before allowing script progression.</summary>
*)
{endregion}
METHOD PROTECTED ProcessAssertions
VAR_INPUT
    Enable : BOOL; //! Enables checking during the active Test phase.
END_VAR
FProgress(Enable := Enable,
    State := State,
    IN := FProgressMatches);
FEvidence(Enable := Enable,
    State := State,
    IN := FEvidenceMatches);
IF Enable THEN
    FStepChecked := TRUE;
END_IF;
END_METHOD

{region 'Documentation'}
(*!
<summary>No Preparation phase is required for this isolated lifecycle test.</summary>
*)
{endregion}
METHOD PROTECTED ProcessPreparations
VAR_INPUT
    // SA0033: Required hook; the test has no Preparation phase.
    {attribute 'analysis' := '-33'}
    Enable : BOOL; //! No preparation action is performed in either phase.
END_VAR
END_METHOD

{region 'Documentation'}
(*!
<summary>Restarts the script and resets its checking Assertions.</summary>
*)
{endregion}
METHOD PROTECTED ProcessReset
FStep := Setup;
FStepChecked := FALSE;
FProgressMatches := TRUE;
FEvidenceMatches := TRUE;
FProgress.Reset();
FEvidence.Reset();
CompleteReset();
END_METHOD

{region 'Documentation'}
(*!
<summary>Performs one subject call per active cycle and advances only after checking Assertions.</summary>
*)
{endregion}
METHOD PROTECTED ProcessTests
VAR_INPUT
    Enable : BOOL; //! Authorizes scenario progression.
END_VAR
IF NOT Enable THEN
    RETURN;
END_IF;
IF FStepChecked THEN
    FStep := FStep + 1;
    FStepChecked := FALSE;
END_IF;
IF FStep > RepeatAgain THEN
    CompleteTests();
    RETURN;
END_IF;
RunStep();
END_METHOD

{region 'Documentation'}
(*!
<summary>Checks first entry, repeated-request completion, held Idle and a second complete Reset interval.</summary>
*)
{endregion}
METHOD PRIVATE RunStep
VAR
    Config : ST_TestSuiteConfig;
    ExpectedState : E_State;
    Snapshot : ST_TestSuiteStatus;
    Index : UINT;
    ResetTransitions : UINT;
    IdleTransitions : UINT;
END_VAR
CASE FStep OF
    Setup:
        IF NOT FCapture.Initialize(Buffer := FEvents,
            FifoControl := FCaptureFifo,
            Status := FCaptureStatus) THEN
            Error(Message := 'Mock Reset capture initialization failed.');
            RETURN;
        END_IF;
        FSubject.BindPublisher(Publisher := FCapture);
        IF NOT FSubject.Initialize(Parent := FSubjectParent,
            SuiteName := 'RepeatedResetMock',
            Config := Config) THEN
            Error(Message := 'Mock Reset subject initialization failed.');
            RETURN;
        END_IF;
        ExpectedState := E_State.Uninitialized;

    RequestFirst, RequestAgain:
        IF FSubject.ReserveResetEvents() <> E_EventReservationResult.Accepted THEN
            Error(Message := 'Mock Reset reservation was rejected.');
            RETURN;
        END_IF;
        FSubject.RequestReset();
        ExpectedState := E_State.Reset;

    RepeatFirst, RepeatAgain:
        FSubject.RequestReset();
        ExpectedState := E_State.Idle;

    HoldIdle:
        ExpectedState := E_State.Idle;
ELSE
    Error(Message := 'Unexpected mock Reset test step.');
    RETURN;
END_CASE;

FSubject();
Snapshot := FSubject.Status;
FProgressMatches := (FSubject.State = ExpectedState)
    AND (Snapshot.Execution.State = ExpectedState)
    AND (FSubject.Result = E_Result.NotEvaluated)
    AND (Snapshot.Execution.Result = E_Result.NotEvaluated)
    AND NOT FSubject.HasError AND NOT Snapshot.Execution.Error
    AND (FSubject.IsReady = (ExpectedState = E_State.Idle))
    AND (Snapshot.Execution.Ready = (ExpectedState = E_State.Idle))
    AND NOT FSubject.IsComplete AND NOT Snapshot.Execution.Completed;
FEvidenceMatches := (FCaptureStatus.LostEventCount = 0)
    AND (Snapshot.TestCaseCountTotal = 0)
    AND (Snapshot.TestCaseCountIdle = 0)
    AND (Snapshot.TestCaseCountRunning = 0)
    AND (Snapshot.TestCaseCountCompleted = 0)
    AND (Snapshot.TestCaseCountError = 0);

IF (FStep = RepeatFirst) OR (FStep = RepeatAgain) THEN
    IF NOT FSubject.FreeReservedEvents() THEN
        FEvidenceMatches := FALSE;
    END_IF;
    FEvidenceMatches := FEvidenceMatches AND (FSubject.ReservedEntryCount = 0)
        AND (FCapture.ReservedEntryCount = 0);
END_IF;
IF FStep = RepeatAgain THEN
    FOR Index := 1 TO CaptureLength DO
        IF (FEvents[Index].SequenceId <> 0)
            AND (FEvents[Index].Name = FSubject.Name)
            AND (FEvents[Index].EventType = E_EventType.StateTransition) THEN
            IF FEvents[Index].State = E_State.Reset THEN
                ResetTransitions := ResetTransitions + 1;
            ELSIF FEvents[Index].State = E_State.Idle THEN
                IdleTransitions := IdleTransitions + 1;
            END_IF;
        END_IF;
    END_FOR;
    FEvidenceMatches := FEvidenceMatches AND (ResetTransitions = 2)
        AND (IdleTransitions = 2);
END_IF;
END_METHOD

END_FUNCTION_BLOCK

// ---- SelfTests/TestCases/TestSuite_TestSuiteLifecycle/Helper/TestSuiteMockProbe.TcPOU
{region 'Documentation'}
(*!
<summary>Binds an isolated publisher before initialization; all mock lifecycle processing remains inherited.</summary>
*)
{endregion}
FUNCTION_BLOCK TestSuiteMockProbe EXTENDS TestSuiteMock

SUPER^();

{region 'Documentation'}
(*!
<summary>Binds the local capture before the first Initialize without modifying the global publisher.</summary>
*)
{endregion}
METHOD PUBLIC BindPublisher
VAR_INPUT
    Publisher : I_EventPublisher; //! Nonzero borrowed capture retained for the subject lifetime.
END_VAR
FEventPublisher := Publisher;
END_METHOD

END_FUNCTION_BLOCK

// ---- SelfTests/TestSuites/TestSuite_RunControlLifecycle.TcPOU
{region 'Documentation'}
(*!
<summary>Groups isolated RunControlBase owner scenarios; the application's real root and publisher remain unchanged.</summary>
*)
{endregion}
FUNCTION_BLOCK TestSuite_RunControlLifecycle EXTENDS TestSuiteBase
VAR
    FInitialization : Test_RunControlInitialization;
    FTaskMapping : Test_RunControlTaskMapping;
    FTestCases : ARRAY[1..TestCaseCapacity] OF I_TestCase;
    FNormalRepeat : Test_RunControlNormalLifecycle;
    FMixedRepeat : Test_RunControlNormalLifecycle;
    FRequests : Test_RunControlRequests;
    FRealComposition : Test_RunControlRealComposition;
    FResetError : Test_RunControlExceptionalLifecycle;
    FResetTimeout : Test_RunControlExceptionalLifecycle;
    FResetErrorTimeout : Test_RunControlExceptionalLifecycle;
    FChildError : Test_RunControlExceptionalLifecycle;
    FUnexpectedChildAbort : Test_RunControlExceptionalLifecycle;
    FExecutionError : Test_RunControlExceptionalLifecycle;
    FExecutionTimeout : Test_RunControlExceptionalLifecycle;
    FAbort : Test_RunControlExceptionalLifecycle;
    FAbortError : Test_RunControlExceptionalLifecycle;
    FAbortTimeout : Test_RunControlExceptionalLifecycle;
    FAbortErrorTimeout : Test_RunControlExceptionalLifecycle;
    FZeroDelay : Test_RunControlCompletion;
    FDefaultDelay : Test_RunControlCompletion;
    FInvalidTime : Test_RunControlCompletion;
    FLateResetChildren : Test_RunControlCompletion;
END_VAR
VAR CONSTANT
    TestCaseCapacity : UINT := 21;
END_VAR

SUPER^();

{region 'Documentation'}
(*!
<summary>Initializes and registers the local root scenarios for serial execution.</summary>
*)
{endregion}
METHOD PROTECTED Configure
VAR_IN_OUT
    // SA0167: Borrowed owner builder; no temporary instance is created.
    {attribute 'analysis' := '-167'}
    Builder : TestSuiteConfigurationBuilder; //! Borrowed owner configuration builder used only during this Configure call; register this owner's concrete children.
END_VAR
VAR
    TestConfig : ST_TestCaseConfig;
END_VAR
Builder.Initialize(Mode := E_OrchestrationMode.Serial,
    TestCases := FTestCases);
FInitialization.Initialize(Parent := THIS^,
    TestName := 'Initialization',
    Config := TestConfig);
Builder.Register(TestCase := FInitialization);
FTaskMapping.Initialize(Parent := THIS^,
    TestName := 'TaskMapping',
    Config := TestConfig);
Builder.Register(TestCase := FTaskMapping);

FNormalRepeat.Initialize(Parent := THIS^,
    TestName := 'NormalRepeat',
    Config := TestConfig);
Builder.Register(TestCase := FNormalRepeat);
FMixedRepeat.Initialize(Parent := THIS^,
    TestName := 'MixedRepeat',
    Config := TestConfig);
Builder.Register(TestCase := FMixedRepeat);
FRequests.Initialize(Parent := THIS^,
    TestName := 'Requests',
    Config := TestConfig);
Builder.Register(TestCase := FRequests);

FResetError.Initialize(Parent := THIS^,
    TestName := 'ResetError',
    Config := TestConfig);
Builder.Register(TestCase := FResetError);
FResetTimeout.Initialize(Parent := THIS^,
    TestName := 'ResetTimeout',
    Config := TestConfig);
Builder.Register(TestCase := FResetTimeout);
FResetErrorTimeout.Initialize(Parent := THIS^,
    TestName := 'ResetErrorTimeout',
    Config := TestConfig);
Builder.Register(TestCase := FResetErrorTimeout);
FChildError.Initialize(Parent := THIS^,
    TestName := 'ChildError',
    Config := TestConfig);
Builder.Register(TestCase := FChildError);
FUnexpectedChildAbort.Initialize(Parent := THIS^,
    TestName := 'UnexpectedChildAbort',
    Config := TestConfig);
Builder.Register(TestCase := FUnexpectedChildAbort);
FExecutionError.Initialize(Parent := THIS^,
    TestName := 'ExecutionError',
    Config := TestConfig);
Builder.Register(TestCase := FExecutionError);
FExecutionTimeout.Initialize(Parent := THIS^,
    TestName := 'ExecutionTimeout',
    Config := TestConfig);
Builder.Register(TestCase := FExecutionTimeout);
FAbort.Initialize(Parent := THIS^,
    TestName := 'Abort',
    Config := TestConfig);
Builder.Register(TestCase := FAbort);
FAbortError.Initialize(Parent := THIS^,
    TestName := 'AbortError',
    Config := TestConfig);
Builder.Register(TestCase := FAbortError);
FAbortTimeout.Initialize(Parent := THIS^,
    TestName := 'AbortTimeout',
    Config := TestConfig);
Builder.Register(TestCase := FAbortTimeout);
FAbortErrorTimeout.Initialize(Parent := THIS^,
    TestName := 'AbortErrorTimeout',
    Config := TestConfig);
Builder.Register(TestCase := FAbortErrorTimeout);

FZeroDelay.Initialize(Parent := THIS^,
    TestName := 'ZeroDelay',
    Config := TestConfig);
Builder.Register(TestCase := FZeroDelay);
FDefaultDelay.Initialize(Parent := THIS^,
    TestName := 'DefaultDelay',
    Config := TestConfig);
Builder.Register(TestCase := FDefaultDelay);
FInvalidTime.Initialize(Parent := THIS^,
    TestName := 'InvalidTime',
    Config := TestConfig);
Builder.Register(TestCase := FInvalidTime);
FLateResetChildren.Initialize(Parent := THIS^,
    TestName := 'LateResetChildren',
    Config := TestConfig);
Builder.Register(TestCase := FLateResetChildren);

FRealComposition.Initialize(Parent := THIS^,
    TestName := 'RealComposition',
    Config := TestConfig);
Builder.Register(TestCase := FRealComposition);
END_METHOD

{region 'Documentation'}
(*!
<summary>Returns a registered scenario using its original array index.</summary>
*)
{endregion}
METHOD PUBLIC GetTestCase : I_TestCase //! Typed child interface at the original array index; zero when no entry is available.
VAR_INPUT
    Index : DINT; //! Original occupied child-array index, rather than an ordinal position.
END_VAR
GetTestCase := 0;
IF (ChildCount = 0) OR (Index < ChildArrayLowerBound)
    OR (DINT_TO_LINT(Index) >= DINT_TO_LINT(ChildArrayLowerBound) + UINT_TO_LINT(ChildCount)) THEN
    RETURN;
END_IF;
GetTestCase := FTestCases[Index];
END_METHOD

{region 'Documentation'}
(*!
<summary>Calls each owned scenario once per initialized Suite cycle.</summary>
*)
{endregion}
METHOD PROTECTED ProcessTestCases
FInitialization();
FTaskMapping();

FNormalRepeat(FirstChildResult := E_Result.Passed);
FMixedRepeat(FirstChildResult := E_Result.Failed);
FRequests();

FResetError(Scenario := E_RunControlLifecycleScenario.ResetError);
FResetTimeout(Scenario := E_RunControlLifecycleScenario.ResetTimeout);
FResetErrorTimeout(Scenario := E_RunControlLifecycleScenario.ResetErrorTimeout);
FChildError(Scenario := E_RunControlLifecycleScenario.ChildError);
FUnexpectedChildAbort(Scenario := E_RunControlLifecycleScenario.UnexpectedChildAbort);
FExecutionError(Scenario := E_RunControlLifecycleScenario.ExecutionError);
FExecutionTimeout(Scenario := E_RunControlLifecycleScenario.ExecutionTimeout);
FAbort(Scenario := E_RunControlLifecycleScenario.Abort);
FAbortError(Scenario := E_RunControlLifecycleScenario.AbortError);
FAbortTimeout(Scenario := E_RunControlLifecycleScenario.AbortTimeout);
FAbortErrorTimeout(Scenario := E_RunControlLifecycleScenario.AbortErrorTimeout);

FZeroDelay(Scenario := E_RunControlCompletionScenario.ZeroDelay);
FDefaultDelay(Scenario := E_RunControlCompletionScenario.DefaultDelay);
FInvalidTime(Scenario := E_RunControlCompletionScenario.InvalidTime);
FLateResetChildren(Scenario := E_RunControlCompletionScenario.LateResetChildren);
FRealComposition();
END_METHOD

END_FUNCTION_BLOCK

// ---- SelfTests/TestCases/TestSuite_RunControlLifecycle/Test_RunControlInitialization.TcPOU
{region 'Documentation'}
(*!
<summary>Checks root initialization, collection handover, automatic Startup Reset and rejected setup.</summary>
<description>
Each Test state is one setup attempt followed by two subject calls. Valid setup comes first
and last; rejected startup configurations must not reuse a previously valid collection.
Initialize must clear previously queued method requests and queue only one Startup Reset
after success. Configure and helper initialization are observed separately from FB execution.
The matched administrative and publisher views refer to one local Event Buffer. A missing
administrative view is injected only for its dedicated rejection scenario. Local ControlData
is overwritten with stale Name/Status before each call to verify the base refreshes it even
when setup is invalid. Checking Assertions retain failures and use the outer publisher.
</description>
*)
{endregion}
FUNCTION_BLOCK Test_RunControlInitialization EXTENDS TestCaseBase
VAR
    FControl : ST_RunControl;
    FSubject : RunControlLifecycleProbe;
    FHelper : SuiteOrchestratorDouble;
    FCapture : EventBuffer;
    FEvents : ARRAY[1..CaptureLength] OF ST_Event;
    FCaptureFifo : ST_FifoStatus;
    FCaptureStatus : ST_EventBufferStatus;
    FFixtureValid : BOOL;
    FAttempt : INT := FirstValidSetup;
    FAttemptStarted : BOOL;
    FChecked : BOOL;
    FPassiveCalls : UINT;
    FExpectedInitialized : BOOL;
    FInitialSequence : UDINT;
    FInitialization : AssertTrue;
    FInitializationMatches : BOOL;
    FConfigureOrder : AssertTrue;
    FConfigureOrderMatches : BOOL;
    FCollection : AssertTrue;
    FCollectionMatches : BOOL;
    FPassiveState : AssertTrue;
    FPassiveStateMatches : BOOL;
    FDiagnostic : AssertTrue;
    FDiagnosticMatches : BOOL;
    FDispatch : AssertTrue;
    FDispatchMatches : BOOL;
    FCaptureIntegrity : AssertTrue;
END_VAR
VAR CONSTANT
    CaptureLength : UINT := 32;
    PassiveCallCount : UINT := 2;
    FirstValidSetup : INT := 1;
    EmptyName : INT := 2;
    InvalidDepth : INT := 3;
    InvalidCharacter : INT := 4;
    OverlengthName : INT := 5;
    MissingBuffer : INT := 6;
    NoRegistration : INT := 7;
    UninitializedChild : INT := 8;
    ZeroExecutionTimeout : INT := 9;
    ZeroResetTimeout : INT := 10;
    ZeroAbortTimeout : INT := 11;
    RejectedHelper : INT := 12;
    FinalValidSetup : INT := 13;
    AttemptCount : INT := 13;
END_VAR

SUPER^();

{region 'Documentation'}
(*!
<summary>Contributes only the checking Assertions, not the intentionally controlled subject results.</summary>
*)
{endregion}
METHOD PROTECTED AggregateResults
VAR_INPUT
    Aggregator : I_ResultAggregator; //! Borrowed result sink owned by the outer Test Case; add this test's checking Assertions without resetting or retaining the sink.
END_VAR
Aggregator.AddProvider(Provider := FInitialization);
Aggregator.AddProvider(Provider := FConfigureOrder);
Aggregator.AddProvider(Provider := FCollection);
Aggregator.AddProvider(Provider := FPassiveState);
Aggregator.AddProvider(Provider := FDiagnostic);
Aggregator.AddProvider(Provider := FDispatch);
Aggregator.AddProvider(Provider := FCaptureIntegrity);
END_METHOD

{region 'Documentation'}
(*!
<summary>Changes one setup condition and records initialization evidence before cyclic subject execution.</summary>
*)
{endregion}
METHOD PRIVATE BeginAttempt
VAR
    Config : ST_RunConfig;
    BufferService : I_EventBuffer;
    RootName : STRING(2 * GVL_Constants.NameLength + 1);
    Initialized : BOOL;
    ExpectedConfigured : BOOL;
    ExpectedHelper : BOOL;
    Index : UINT;
    FirstChild : I_Orchestratable;
    LastChild : I_Orchestratable;
    SubjectCollection : I_OrchestratableCollection;
    Publisher : I_EventPublisher;
    SubjectStatus : ST_RunControlStatus;
    FirstSharedChild : I_Orchestratable;
    LastSharedChild : I_Orchestratable;
    BelowRangeChild : I_Orchestratable;
    UnusedChild : I_Orchestratable;
    UnusedTypedChild : I_TestSuite;
END_VAR
FFixtureValid := FCapture.Initialize(Buffer := FEvents,
    FifoControl := FCaptureFifo,
    Status := FCaptureStatus);
IF NOT FFixtureValid THEN
    Error(Message := 'Run Control initialization capture could not be initialized.');
    RETURN;
END_IF;
BufferService := FCapture;
RootName := 'RootSubject';
CASE FAttempt OF
    EmptyName:
        RootName := '';
    InvalidDepth:
        RootName := 'Invalid.Root';
    InvalidCharacter:
        RootName := 'Invalid Root';
    OverlengthName:
        FOR Index := 1 TO GVL_Constants.NameLength DO
            RootName := CONCAT(RootName, 'x');
        END_FOR;
    MissingBuffer:
        BufferService := 0;
    ZeroExecutionTimeout:
        Config.Timeout := T#0s;
    ZeroResetTimeout:
        Config.ResetTimeout := T#0s;
    ZeroAbortTimeout:
        Config.AbortTimeout := T#0s;
ELSE
    // Remaining attempts vary the concrete setup or helper, not these external inputs.
END_CASE;
FExpectedInitialized := (FAttempt = FirstValidSetup) OR (FAttempt = FinalValidSetup);
ExpectedConfigured := FExpectedInitialized OR (FAttempt >= NoRegistration);
ExpectedHelper := ExpectedConfigured AND (FAttempt <> NoRegistration);
FHelper.BeginScenario(AcceptInitialization := FAttempt <> RejectedHelper);
FSubject.Bind(Publisher := FCapture,
    Helper := FHelper,
    Config := Config,
    RegisterChildren := FAttempt <> NoRegistration,
    IncludeUninitializedChild := FAttempt = UninitializedChild);
FSubject.RequestStart();
FSubject.RequestAbort();
FSubject.RequestReset();
Initialized := FSubject.Initialize(Name := RootName,
    EventBuffer := BufferService);
Publisher := FCapture;
SubjectStatus := FSubject.Status;
FInitializationMatches := (Initialized = FExpectedInitialized)
    AND (FSubject.IsInitialized = FExpectedInitialized)
    AND (SubjectStatus.Execution.ConfigError <> FExpectedInitialized)
    AND (FSubject.EventPublisher = Publisher);
IF FAttempt = OverlengthName THEN
    FInitializationMatches := FInitializationMatches AND (LEN(FSubject.Name) = GVL_Constants.NameLength);
ELSE
    FInitializationMatches := FInitializationMatches AND (FSubject.Name = RootName);
END_IF;
FConfigureOrderMatches := FSubject.ConfigureCount = BOOL_TO_UINT(ExpectedConfigured);
IF ExpectedConfigured THEN
    FConfigureOrderMatches := FConfigureOrderMatches AND FSubject.ConfigureContextValid;
END_IF;
FCollectionMatches := FHelper.InitializeCount = BOOL_TO_UINT(ExpectedHelper);
IF ExpectedHelper THEN
    SubjectCollection := FSubject;
    FCollectionMatches := FCollectionMatches
        AND (FHelper.Collection = SubjectCollection)
        AND (FHelper.FirstIndex = 4) AND (FHelper.LastIndex = 6) AND (FHelper.ChildCount = 2)
        AND (FHelper.FirstChild <> 0) AND (FHelper.LastChild <> 0)
        AND (FHelper.FirstChild <> FHelper.LastChild)
        AND (FHelper.OwnerName = FSubject.Name) AND (FHelper.ResourceName = 'Fixture');
END_IF;
FirstSharedChild := FSubject.GetChild(Index := 4);
LastSharedChild := FSubject.GetChild(Index := 5);
BelowRangeChild := FSubject.GetChild(Index := 3);
UnusedChild := FSubject.GetChild(Index := 6);
UnusedTypedChild := FSubject.GetTestSuite(Index := 6);
IF FExpectedInitialized THEN
    FirstChild := FSubject.GetTestSuite(Index := 4);
    LastChild := FSubject.GetTestSuite(Index := 5);
    FCollectionMatches := FCollectionMatches
        AND (FSubject.ChildCount = 2)
        AND (FSubject.ChildArrayLowerBound = 4) AND (FSubject.ChildArrayUpperBound = 6)
        AND (FirstSharedChild = FirstChild)
        AND (LastSharedChild = LastChild)
        AND (FHelper.FirstChild = FirstChild) AND (FHelper.LastChild = LastChild)
        AND (BelowRangeChild = 0) AND (UnusedChild = 0)
        AND (UnusedTypedChild = 0)
        AND (FSubject.Name = 'RootSubject');
ELSE
    FirstChild := FSubject.GetTestSuite(Index := 4);
    FCollectionMatches := FCollectionMatches
        AND (FSubject.ChildCount = 0)
        AND (FSubject.ChildArrayLowerBound = 0) AND (FSubject.ChildArrayUpperBound = 0)
        AND (FirstSharedChild = 0) AND (FirstChild = 0);
END_IF;
FInitialSequence := FCaptureStatus.SequenceId;
IF FExpectedInitialized THEN
    FDiagnosticMatches := FInitialSequence = 0;
ELSE
    FDiagnosticMatches := (FInitialSequence = 1)
        AND (FEvents[1].EventType = E_EventType.Framework)
        AND (FEvents[1].Severity = E_EventSeverity.Error)
        AND (FEvents[1].State = E_State.Uninitialized)
        AND (FEvents[1].Name = FSubject.Name);
END_IF;
FPassiveStateMatches := (FSubject.State = E_State.Uninitialized) AND NOT FSubject.IsReady;
FDispatchMatches := (FHelper.ExecuteCount = 0) AND (FSubject.ChildCallCount = 0);
FPassiveCalls := 0;
FAttemptStarted := TRUE;
END_METHOD

{region 'Documentation'}
(*!
<summary>Initializes the checking Assertions; the scenario explicitly initializes its isolated subject.</summary>
*)
{endregion}
METHOD PROTECTED Configure
FPreparationStateCount := 0;
FTestStateCount := AttemptCount;
FInitialization.Initialize(Parent := THIS^,
    AssertionName := 'Initialization');
FConfigureOrder.Initialize(Parent := THIS^,
    AssertionName := 'ConfigureOrder');
FCollection.Initialize(Parent := THIS^,
    AssertionName := 'Collection');
FPassiveState.Initialize(Parent := THIS^,
    AssertionName := 'PassiveState');
FDiagnostic.Initialize(Parent := THIS^,
    AssertionName := 'Diagnostic');
FDispatch.Initialize(Parent := THIS^,
    AssertionName := 'Dispatch');
FCaptureIntegrity.Initialize(Parent := THIS^,
    AssertionName := 'CaptureIntegrity');
END_METHOD

{region 'Documentation'}
(*!
<summary>No asynchronous test resource remains to stop.</summary>
*)
{endregion}
METHOD PROTECTED ProcessAbort
VAR_INPUT
    Enable : BOOL; //! Phase permission supplied by the owning Test Case; FALSE does not authorize progression, while observation may continue.
END_VAR
IF Enable THEN
    CompleteAbort();
END_IF;
END_METHOD

{region 'Documentation'}
(*!
<summary>Latches each setup after two calls: successful startup consumes Reset once; rejected setup stays passive.</summary>
*)
{endregion}
METHOD PROTECTED ProcessAssertions
VAR_INPUT
    Enable : BOOL; //! Phase permission supplied by the owning Test Case; FALSE does not authorize progression, while observation may continue.
END_VAR
VAR
    Evaluate : BOOL;
END_VAR
Evaluate := Enable AND (FPassiveCalls >= PassiveCallCount);
FInitialization(Enable := Evaluate,
    State := State,
    IN := FInitializationMatches);
FConfigureOrder(Enable := Evaluate,
    State := State,
    IN := FConfigureOrderMatches);
FCollection(Enable := Evaluate,
    State := State,
    IN := FCollectionMatches);
FPassiveState(Enable := Evaluate,
    State := State,
    IN := FPassiveStateMatches);
FDiagnostic(Enable := Evaluate,
    State := State,
    IN := FDiagnosticMatches);
FDispatch(Enable := Evaluate,
    State := State,
    IN := FDispatchMatches);
FCaptureIntegrity(Enable := Evaluate,
    State := State,
    IN := FCaptureStatus.LostEventCount = 0);
IF Evaluate THEN
    FChecked := TRUE;
END_IF;
END_METHOD

{region 'Documentation'}
(*!
<summary>No resource Preparation is required for this controlled owner scenario.</summary>
*)
{endregion}
METHOD PROTECTED ProcessPreparations
VAR_INPUT
    // SA0033: Required override; the scenario has no Preparation phase.
    {attribute 'analysis' := '-33'}
    Enable : BOOL; //! Phase permission supplied by the owning Test Case; FALSE does not authorize progression, while observation may continue.
END_VAR
END_METHOD

{region 'Documentation'}
(*!
<summary>Restarts the test script and clears checking Assertions; subject setup belongs to the next test attempt.</summary>
*)
{endregion}
METHOD PROTECTED ProcessReset
FAttempt := FirstValidSetup;
FAttemptStarted := FALSE;
FChecked := FALSE;
FPassiveCalls := 0;
FInitialization.Reset();
FConfigureOrder.Reset();
FCollection.Reset();
FPassiveState.Reset();
FDiagnostic.Reset();
FDispatch.Reset();
FCaptureIntegrity.Reset();
CompleteReset();
END_METHOD

{region 'Documentation'}
(*!
<summary>Advances the explicit test script with at most one subject FB call per active PLC cycle.</summary>
*)
{endregion}
METHOD PROTECTED ProcessTests
VAR_INPUT
    Enable : BOOL; //! Phase permission supplied by the owning Test Case; FALSE does not authorize progression, while observation may continue.
END_VAR
IF NOT Enable THEN
    RETURN;
END_IF;
IF FChecked THEN
    IF FAttempt = AttemptCount THEN
        CompleteTests();
        RETURN;
    END_IF;
    FAttempt := FAttempt + 1;
    FAttemptStarted := FALSE;
    FChecked := FALSE;
    NextTestState();
END_IF;
IF NOT FAttemptStarted THEN
    BeginAttempt();
    IF NOT FFixtureValid THEN
        RETURN;
    END_IF;
END_IF;
// Deliberately stale public data must be replaced even after rejected initialization.
FControl.Name := 'Stale';
FControl.Status.Execution.State := E_State.Completed;
FControl.Status.Execution.Ready := TRUE;
FSubject(ControlData := FControl);
FPassiveCalls := FPassiveCalls + 1;
FPassiveStateMatches := FPassiveStateMatches
    AND NOT FSubject.IsReady AND (FSubject.Result = E_Result.NotEvaluated)
    AND (FControl.Name = FSubject.Name)
    AND (FControl.Status.Execution.State = FSubject.State)
    AND (FControl.Status.Execution.Result = FSubject.Result)
    AND (FControl.Status.Execution.Ready = FSubject.IsReady)
    AND (FControl.Status.Execution.ConfigError <> FExpectedInitialized);
IF FExpectedInitialized THEN
    FPassiveStateMatches := FPassiveStateMatches AND (FSubject.State = E_State.Reset);
    FDispatchMatches := FDispatchMatches
        AND (FHelper.ExecuteCount = FPassiveCalls)
        AND (FSubject.ChildCallCount = FPassiveCalls)
        AND FSubject.ChildBodyCallsMatch
        AND (FHelper.CurrentTask = E_OrchestratorTask.Reset);
    FDiagnosticMatches := FDiagnosticMatches
        AND (FCaptureStatus.SequenceId = 2)
        AND (FEvents[1].EventType = E_EventType.Trigger)
        AND (FEvents[1].State = E_State.Uninitialized)
        AND (FEvents[2].EventType = E_EventType.StateTransition)
        AND (FEvents[2].State = E_State.Reset);
ELSE
    FPassiveStateMatches := FPassiveStateMatches AND (FSubject.State = E_State.Uninitialized);
    FDispatchMatches := FDispatchMatches
        AND (FHelper.ExecuteCount = 0) AND (FSubject.ChildCallCount = 0);
    FDiagnosticMatches := FDiagnosticMatches AND (FCaptureStatus.SequenceId = FInitialSequence);
END_IF;
END_METHOD

END_FUNCTION_BLOCK

// ---- SelfTests/TestCases/TestSuite_RunControlLifecycle/Helper/RunControlLifecycleProbe.TcPOU
{region 'Documentation'}
(*!
<summary>Thin RunControlBase subject with a typed child array and isolated dependencies.</summary>
<description>
Bind is called before Initialize. Production initialization, sequencing, aggregation and
publication remain inherited. Configure records its context and builds a small real collection.
The uninitialized-child option uses a separate never-initialized double, not mutated base state.
ProcessTestSuites applies the scenario's child view only after the base has called its helper.
</description>
*)
{endregion}
FUNCTION_BLOCK RunControlLifecycleProbe EXTENDS RunControlBase
VAR
    FChildA : RunControlSuiteDouble;
    FChildB : RunControlSuiteDouble;
    FUninitializedChild : RunControlSuiteDouble;
    FTestSuites : ARRAY[4..6] OF I_TestSuite;
    FChildObservation : ST_OrchestrationObservation;
    FSecondChildObservation : ST_OrchestrationObservation;
    FSelectedConfig : ST_RunConfig;
    FRegisterChildren : BOOL := TRUE;
    FIncludeUninitializedChild : BOOL;
    FConfigureCount : UINT;
    FConfigureContextValid : BOOL;
    FChildCallCount : UINT;
    FForceInvalidCompletionTime : BOOL;
END_VAR

SUPER^(ControlData := ControlData);

{region 'Documentation'}
(*!
<summary>Binds isolated dependencies before Initialize and selects the concrete setup to exercise.</summary>
*)
{endregion}
METHOD PUBLIC Bind
VAR_INPUT
    Publisher : I_EventPublisher; //! Nonzero isolated event publisher retained before subject initialization; keep it alive through all subject use.
    Helper : I_Orchestrator; //! Nonzero injected orchestration helper retained before owner initialization; keep it alive through subject use.
    Config : ST_RunConfig; //! Run configuration copied for the next owner initialization.
    RegisterChildren : BOOL := TRUE; //! TRUE registers the two controlled children; FALSE exercises empty configuration.
    IncludeUninitializedChild : BOOL := FALSE; //! TRUE leaves a registered controlled child uninitialized to exercise rejection.
END_VAR
FEventPublisher := Publisher;
FOrchestrator := Helper;
FSelectedConfig := Config;
FRegisterChildren := RegisterChildren;
FIncludeUninitializedChild := IncludeUninitializedChild;
FForceInvalidCompletionTime := FALSE;
FConfigureCount := 0;
FChildCallCount := 0;
FConfigureContextValid := FALSE;
FChildObservation.State := E_State.Uninitialized;
FChildObservation.Result := E_Result.NotEvaluated;
FChildObservation.Ready := FALSE;
FChildObservation.Complete := FALSE;
FSecondChildObservation := FChildObservation;
END_METHOD

{region 'Documentation'}
(*!
<summary>Both concrete child bodies have executed exactly once per ProcessTestSuites invocation.</summary>
*)
{endregion}
{attribute 'monitoring' := 'call'}
PROPERTY PUBLIC ChildBodyCallsMatch : BOOL //! Both concrete child bodies have executed exactly once per ProcessTestSuites invocation.
GET
VAR
    FirstCalls : ST_OrchestrationCalls;
    SecondCalls : ST_OrchestrationCalls;
END_VAR
FirstCalls := FChildA.Calls;
SecondCalls := FChildB.Calls;
ChildBodyCallsMatch := (FirstCalls.BodyCount = FChildCallCount) AND (SecondCalls.BodyCount = FChildCallCount);
END_GET
END_PROPERTY

{region 'Documentation'}
(*!
<summary>Number of ProcessTestSuites invocations since binding.</summary>
*)
{endregion}
{attribute 'monitoring' := 'call'}
PROPERTY PUBLIC ChildCallCount : UINT //! Number of ProcessTestSuites invocations since binding.
GET
ChildCallCount := FChildCallCount;
END_GET
END_PROPERTY

{region 'Documentation'}
(*!
<summary>Registers two controlled typed children in a shifted array with spare capacity; records base context.</summary>
*)
{endregion}
METHOD PROTECTED Configure
VAR_IN_OUT
    // SA0167: Borrowed setup builder; no temporary instance is created.
    {attribute 'analysis' := '-167'}
    Builder : RunControlConfigurationBuilder; //! Borrowed owner configuration builder used only during this Configure call; register this owner's concrete children.
END_VAR
FConfig := FSelectedConfig;
FResourceName := 'Fixture';
FConfigureCount := FConfigureCount + 1;
FConfigureContextValid := (State = E_State.Uninitialized) AND NOT IsInitialized AND (Name <> '');
Builder.Initialize(Mode := E_OrchestrationMode.Serial,
    TestSuites := FTestSuites);
FChildA.Initialize(Name := CONCAT(Name, '.ChildA'),
    Slot := 0);
FChildB.Initialize(Name := CONCAT(Name, '.ChildB'),
    Slot := 0);
IF NOT FRegisterChildren THEN
    RETURN;
END_IF;
Builder.Register(TestSuite := FChildA);
IF FIncludeUninitializedChild THEN
    Builder.Register(TestSuite := FUninitializedChild);
ELSE
    Builder.Register(TestSuite := FChildB);
END_IF;
END_METHOD

{region 'Documentation'}
(*!
<summary>Configure saw the new identity before successful initialization.</summary>
*)
{endregion}
{attribute 'monitoring' := 'call'}
PROPERTY PUBLIC ConfigureContextValid : BOOL //! Configure saw the new identity before successful initialization.
GET
ConfigureContextValid := FConfigureContextValid;
END_GET
END_PROPERTY

{region 'Documentation'}
(*!
<summary>Number of Configure calls since binding.</summary>
*)
{endregion}
{attribute 'monitoring' := 'call'}
PROPERTY PUBLIC ConfigureCount : UINT //! Number of Configure calls since binding.
GET
ConfigureCount := FConfigureCount;
END_GET
END_PROPERTY

{region 'Documentation'}
(*!
<summary>Returns the recorded calls of a registered controlled child; unknown indices return an empty observation.</summary>
*)
{endregion}
METHOD PUBLIC GetChildCalls : ST_OrchestrationCalls //! Retained call trace for the selected child; an empty trace for an unknown index or empty collection.
VAR_INPUT
    Index : DINT; //! Original occupied child-array index; unknown indices return an empty trace.
END_VAR
VAR
    EmptyCalls : ST_OrchestrationCalls;
END_VAR
GetChildCalls := EmptyCalls;
IF ChildCount = 0 THEN
    RETURN;
END_IF;
IF Index = ChildArrayLowerBound THEN
    GetChildCalls := FChildA.Calls;
ELSIF (ChildCount > 1) AND (Index = ChildArrayLowerBound + 1) THEN
    GetChildCalls := FChildB.Calls;
END_IF;
END_METHOD

{region 'Documentation'}
(*!
<summary>Returns the registered typed entry by actual array index; lookup never executes a child.</summary>
*)
{endregion}
METHOD PUBLIC GetTestSuite : I_TestSuite //! Typed Suite interface at the original array index; zero when no entry is available.
VAR_INPUT
    Index : DINT; //! Original occupied child-array index, rather than an ordinal position.
END_VAR
GetTestSuite := 0;
IF (ChildCount = 0) OR (Index < ChildArrayLowerBound)
    OR (DINT_TO_LINT(Index) >= DINT_TO_LINT(ChildArrayLowerBound) + UINT_TO_LINT(ChildCount)) THEN
    RETURN;
END_IF;
GetTestSuite := FTestSuites[Index];
END_METHOD

{region 'Documentation'}
(*!
<summary>Overrides only completion validity; the real timer and all elapsed-time calculations remain unchanged.</summary>
*)
{endregion}
{attribute 'monitoring' := 'call'}
PROPERTY PROTECTED IsCompletionTimeValid : BOOL //! Overrides only completion validity; the real timer and all elapsed-time calculations remain unchanged.
GET
IsCompletionTimeValid := SUPER^.IsCompletionTimeValid AND NOT FForceInvalidCompletionTime;
END_GET
END_PROPERTY

{region 'Documentation'}
(*!
<summary>Applies the next scripted observation after the helper; counts calls without replacing owner processing.</summary>
*)
{endregion}
METHOD PROTECTED ProcessTestSuites
FChildA(ObservationInput := FChildObservation);
FChildB(ObservationInput := FSecondChildObservation);
FChildCallCount := FChildCallCount + 1;
END_METHOD

{region 'Documentation'}
(*!
<summary>Selects the next child snapshot; it becomes visible only in ProcessTestSuites, after helper execution.</summary>
*)
{endregion}
METHOD PUBLIC SetChildObservation
VAR_INPUT
    Observation : ST_OrchestrationObservation; //! Scripted view copied to both children for acceptance on their next concrete body calls.
END_VAR
FChildObservation := Observation;
FSecondChildObservation := Observation;
END_METHOD

{region 'Documentation'}
(*!
<summary>Supplies independent next snapshots; each child accepts its view only when the Run-Control calls its body.</summary>
*)
{endregion}
METHOD PUBLIC SetChildObservations
VAR_INPUT
    FirstChild : ST_OrchestrationObservation; //! Scripted view for the first child, accepted on its next concrete body call.
    SecondChild : ST_OrchestrationObservation; //! Scripted view for the second child, accepted on its next concrete body call.
END_VAR
FChildObservation := FirstChild;
FSecondChildObservation := SecondChild;
END_METHOD

{region 'Documentation'}
(*!
<summary>Controls the test-only validity observation; Bind restores the default real-clock behavior.</summary>
*)
{endregion}
METHOD PUBLIC SetInvalidCompletionTime
VAR_INPUT
    Invalid : BOOL; //! TRUE forces the completion-validity seam to FALSE without replacing clock or elapsed-time calculations.
END_VAR
FForceInvalidCompletionTime := Invalid;
END_METHOD

END_FUNCTION_BLOCK

// ---- SelfTests/TestCases/TestSuite_RunControlLifecycle/Helper/RunControlSuiteDouble.TcPOU
{region 'Documentation'}
(*!
<summary>Adds the typed Test Suite status to the existing scripted child boundary; requests remain observation-only.</summary>
*)
{endregion}
FUNCTION_BLOCK RunControlSuiteDouble EXTENDS OrchestrationChildDouble IMPLEMENTS I_TestSuite

SUPER^(ObservationInput := ObservationInput);

{region 'Documentation'}
(*!
<summary>Projects the scripted child observation into the typed Run-Control-facing status; no lifecycle is copied.</summary>
*)
{endregion}
{attribute 'monitoring' := 'variable'}
PROPERTY PUBLIC Status : ST_TestSuiteStatus //! Projects the scripted child observation into the typed Run-Control-facing status; no lifecycle is copied.
GET
VAR
    Snapshot : ST_TestSuiteStatus;
    View : ST_OrchestrationObservation;
END_VAR
View := Observation;
Snapshot.Execution.State := View.State;
Snapshot.Execution.Result := View.Result;
Snapshot.Execution.Ready := View.Ready;
Snapshot.Execution.Completed := View.Complete;
Snapshot.Execution.Error := View.Result = E_Result.Error;
CASE View.State OF
    E_State.Uninitialized:
        Snapshot.Execution.ExecutionStatus := E_ExecutionStatus.NotReady;
        Snapshot.Execution.Uninitialized := TRUE;
    E_State.Reset:
        Snapshot.Execution.ExecutionStatus := E_ExecutionStatus.Reset;
    E_State.Idle:
        Snapshot.Execution.ExecutionStatus := E_ExecutionStatus.Idle;
    E_State.Starting:
        Snapshot.Execution.ExecutionStatus := E_ExecutionStatus.Starting;
    E_State.Running:
        Snapshot.Execution.ExecutionStatus := E_ExecutionStatus.Running;
        Snapshot.Execution.Running := TRUE;
    E_State.Completing:
        Snapshot.Execution.ExecutionStatus := E_ExecutionStatus.Completing;
    E_State.Completed:
        Snapshot.Execution.ExecutionStatus := E_ExecutionStatus.Completed;
    E_State.Aborting, E_State.AbortingFromError:
        Snapshot.Execution.ExecutionStatus := E_ExecutionStatus.Aborting;
ELSE
    Snapshot.Execution.ExecutionStatus := E_ExecutionStatus.Error;
END_CASE;
Status := Snapshot;
END_GET
END_PROPERTY

END_FUNCTION_BLOCK

// ---- SelfTests/TestCases/TestSuite_RunControlLifecycle/Test_RunControlTaskMapping.TcPOU
{region 'Documentation'}
(*!
<summary>Observes RunControlBase task mapping through the controlled helper, not a copied scheduler.</summary>
<description>
Each Test state performs one subject call. Startup Reset remains pending until the helper
reports completion. Readiness can then change in Idle without another Reset.
A short Start/Abort path covers Execution, Abort, completing-task retention and completed Idle.
It is a mapping probe; request priorities, detailed result payloads and deadlines have their
own scenarios. Child snapshots become visible only through ProcessTestSuites.
The subject uses local ControlData and a local Event Buffer; the outer root is never replaced.
</description>
*)
{endregion}
FUNCTION_BLOCK Test_RunControlTaskMapping EXTENDS TestCaseBase
VAR
    FSubject : RunControlLifecycleProbe;
    FHelper : SuiteOrchestratorDouble;
    FControl : ST_RunControl;
    FCapture : EventBuffer;
    FEvents : ARRAY[1..CaptureLength] OF ST_Event;
    FCaptureFifo : ST_FifoStatus;
    FCaptureStatus : ST_EventBufferStatus;
    FStep : INT := StartupReset;
    FChecked : BOOL;
    FStepExecuted : BOOL;
    FExpectedState : E_State;
    FExpectedTask : E_OrchestratorTask;
    FExpectedReady : BOOL;
    FExpectedTriggers : UINT;
    FTriggerCount : UINT;
    FBeforeFirstCallMatches : BOOL;
    FStateMapping : AssertTrue;
    FReadiness : AssertTrue;
    FDispatch : AssertTrue;
    FPublicStatus : AssertTrue;
    FStartupReset : AssertTrue;
    FCaptureIntegrity : AssertTrue;
END_VAR
VAR CONSTANT
    CaptureLength : UINT := 32;
    StartupReset : INT := 1;
    HoldReset : INT := 2;
    FinishReset : INT := 3;
    ReadyIdle : INT := 4;
    WithdrawReady : INT := 5;
    RestoreReady : INT := 6;
    StartExecution : INT := 7;
    Running : INT := 8;
    AbortRequestStep : INT := 9;
    HoldAbort : INT := 10;
    ObserveAbortedChildren : INT := 11;
    Completing : INT := 12;
    Completed : INT := 13;
    HoldCompleted : INT := 14;
    StepCount : INT := 14;
END_VAR

SUPER^();

{region 'Documentation'}
(*!
<summary>Contributes only the checking Assertions, not the intentionally controlled subject results.</summary>
*)
{endregion}
METHOD PROTECTED AggregateResults
VAR_INPUT
    Aggregator : I_ResultAggregator; //! Borrowed result sink owned by the outer Test Case; add this test's checking Assertions without resetting or retaining the sink.
END_VAR
Aggregator.AddProvider(Provider := FStateMapping);
Aggregator.AddProvider(Provider := FReadiness);
Aggregator.AddProvider(Provider := FDispatch);
Aggregator.AddProvider(Provider := FPublicStatus);
Aggregator.AddProvider(Provider := FStartupReset);
Aggregator.AddProvider(Provider := FCaptureIntegrity);
END_METHOD

{region 'Documentation'}
(*!
<summary>Initializes the checking Assertions; the scenario explicitly initializes its isolated subject.</summary>
*)
{endregion}
METHOD PROTECTED Configure
FPreparationStateCount := 0;
FTestStateCount := StepCount;
FStateMapping.Initialize(Parent := THIS^,
    AssertionName := 'StateMapping');
FReadiness.Initialize(Parent := THIS^,
    AssertionName := 'Readiness');
FDispatch.Initialize(Parent := THIS^,
    AssertionName := 'Dispatch');
FPublicStatus.Initialize(Parent := THIS^,
    AssertionName := 'PublicStatus');
FStartupReset.Initialize(Parent := THIS^,
    AssertionName := 'StartupReset');
FCaptureIntegrity.Initialize(Parent := THIS^,
    AssertionName := 'CaptureIntegrity');
END_METHOD

{region 'Documentation'}
(*!
<summary>No asynchronous test resource remains to stop.</summary>
*)
{endregion}
METHOD PROTECTED ProcessAbort
VAR_INPUT
    Enable : BOOL; //! Phase permission supplied by the owning Test Case; FALSE does not authorize progression, while observation may continue.
END_VAR
IF Enable THEN
    CompleteAbort();
END_IF;
END_METHOD

{region 'Documentation'}
(*!
<summary>Checks every scripted mapping step and latches any deviation across the whole scenario.</summary>
*)
{endregion}
METHOD PROTECTED ProcessAssertions
VAR_INPUT
    Enable : BOOL; //! Phase permission supplied by the owning Test Case; FALSE does not authorize progression, while observation may continue.
END_VAR
VAR
    Evaluate : BOOL;
END_VAR
Evaluate := Enable AND FStepExecuted;
FStateMapping(Enable := Evaluate,
    State := State,
    IN := (FSubject.State = FExpectedState) AND (FHelper.CurrentTask = FExpectedTask)
        AND (FSubject.Result <> E_Result.Error));
FReadiness(Enable := Evaluate,
    State := State,
    IN := FSubject.IsReady = FExpectedReady);
FDispatch(Enable := Evaluate,
    State := State,
    IN := (FHelper.ExecuteCount = INT_TO_UINT(FStep))
        AND (FSubject.ChildCallCount = INT_TO_UINT(FStep))
        AND FSubject.ChildBodyCallsMatch
        AND (FSubject.ConfigureCount = 1) AND (FHelper.InitializeCount = 1));
FPublicStatus(Enable := Evaluate,
    State := State,
    IN := (FControl.Name = 'MappingSubject')
        AND (FControl.Status.Execution.State = FExpectedState)
        AND (FControl.Status.Execution.Ready = FExpectedReady)
        AND (FControl.Status.Execution.Result = FSubject.Result)
        AND NOT FControl.Status.Execution.ConfigError
        AND (FControl.Status.SuiteCountTotal = 2));
FStartupReset(Enable := Evaluate,
    State := State,
    IN := FBeforeFirstCallMatches AND (FTriggerCount = FExpectedTriggers)
        AND (FEvents[1].EventType = E_EventType.Trigger)
        AND (FEvents[1].State = E_State.Uninitialized));
FCaptureIntegrity(Enable := Evaluate,
    State := State,
    IN := FCaptureStatus.LostEventCount = 0);
IF Evaluate THEN
    FChecked := TRUE;
END_IF;
END_METHOD

{region 'Documentation'}
(*!
<summary>No resource Preparation is required for this controlled owner scenario.</summary>
*)
{endregion}
METHOD PROTECTED ProcessPreparations
VAR_INPUT
    // SA0033: Required override; the scenario has no Preparation phase.
    {attribute 'analysis' := '-33'}
    Enable : BOOL; //! Phase permission supplied by the owning Test Case; FALSE does not authorize progression, while observation may continue.
END_VAR
END_METHOD

{region 'Documentation'}
(*!
<summary>Restarts the test script and clears checking Assertions; subject setup belongs to the next test attempt.</summary>
*)
{endregion}
METHOD PROTECTED ProcessReset
FStep := StartupReset;
FChecked := FALSE;
FStepExecuted := FALSE;
FStateMapping.Reset();
FReadiness.Reset();
FDispatch.Reset();
FPublicStatus.Reset();
FStartupReset.Reset();
FCaptureIntegrity.Reset();
CompleteReset();
END_METHOD

{region 'Documentation'}
(*!
<summary>Advances the explicit test script with at most one subject FB call per active PLC cycle.</summary>
*)
{endregion}
METHOD PROTECTED ProcessTests
VAR_INPUT
    Enable : BOOL; //! Phase permission supplied by the owning Test Case; FALSE does not authorize progression, while observation may continue.
END_VAR
VAR
    Config : ST_RunConfig;
    ChildView : ST_OrchestrationObservation;
    Index : UINT;
END_VAR
IF NOT Enable THEN
    RETURN;
END_IF;
IF FChecked THEN
    IF FStep = StepCount THEN
        CompleteTests();
        RETURN;
    END_IF;
    FStep := FStep + 1;
    FChecked := FALSE;
    FStepExecuted := FALSE;
    NextTestState();
END_IF;
IF FStep = StartupReset THEN
    IF NOT FCapture.Initialize(Buffer := FEvents,
        FifoControl := FCaptureFifo,
        Status := FCaptureStatus) THEN
        Error(Message := 'Run Control task-mapping capture could not be initialized.');
        RETURN;
    END_IF;
    Config.CompletionDelay := T#0ms;
    FHelper.BeginScenario();
    FSubject.Bind(Publisher := FCapture,
        Helper := FHelper,
        Config := Config);
    IF NOT FSubject.Initialize(Name := 'MappingSubject',
        EventBuffer := FCapture) THEN
        Error(Message := 'Run Control task-mapping subject could not be initialized.');
        RETURN;
    END_IF;
    FBeforeFirstCallMatches := (FSubject.State = E_State.Uninitialized)
        AND NOT FSubject.IsReady AND (FHelper.ExecuteCount = 0)
        AND (FSubject.ChildCallCount = 0) AND (FCaptureStatus.SequenceId = 0);
END_IF;

FExpectedState := E_State.Idle;
FExpectedTask := E_OrchestratorTask.Idle;
FExpectedReady := FALSE;
FExpectedTriggers := 1;
ChildView.State := E_State.Idle;
ChildView.Ready := TRUE;
FHelper.SetObservation(Ready := FALSE);
CASE FStep OF
    StartupReset, HoldReset:
        FExpectedState := E_State.Reset;
        FExpectedTask := E_OrchestratorTask.Reset;
    FinishReset:
        FHelper.SetObservation(Ready := FALSE,
            ResetFinished := TRUE);
    ReadyIdle, RestoreReady:
        FHelper.SetObservation(Ready := TRUE);
        FExpectedReady := TRUE;
    WithdrawReady:
        FHelper.SetObservation(Ready := FALSE);
    StartExecution:
        FHelper.SetObservation(Ready := TRUE);
        FSubject.RequestStart();
        FExpectedState := E_State.Starting;
        FExpectedTask := E_OrchestratorTask.Execution;
        FExpectedTriggers := 2;
        ChildView.State := E_State.Running;
        ChildView.Ready := FALSE;
    Running:
        FExpectedState := E_State.Running;
        FExpectedTask := E_OrchestratorTask.Execution;
        FExpectedTriggers := 2;
        ChildView.State := E_State.Running;
        ChildView.Ready := FALSE;
    AbortRequestStep, HoldAbort:
        IF FStep = AbortRequestStep THEN
            FSubject.RequestAbort();
        END_IF;
        FExpectedState := E_State.Aborting;
        FExpectedTask := E_OrchestratorTask.Abort;
        FExpectedTriggers := 3;
        ChildView.State := E_State.Running;
        ChildView.Ready := FALSE;
    ObserveAbortedChildren, Completing, Completed, HoldCompleted:
        ChildView.State := E_State.Completed;
        ChildView.Ready := FALSE;
        ChildView.Result := E_Result.Abort;
        ChildView.Complete := TRUE;
        FExpectedTriggers := 3;
        CASE FStep OF
            ObserveAbortedChildren:
                FExpectedState := E_State.Aborting;
                FExpectedTask := E_OrchestratorTask.Abort;
            Completing:
                FHelper.SetObservation(Ready := FALSE,
                    AbortFinished := TRUE);
                FExpectedState := E_State.Completing;
                FExpectedTask := E_OrchestratorTask.Abort;
        ELSE
            FExpectedState := E_State.Completed;
        END_CASE;
END_CASE;
FSubject.SetChildObservation(Observation := ChildView);
FSubject(ControlData := FControl);
FTriggerCount := 0;
FOR Index := 1 TO FCaptureFifo.ElementCount DO
    IF FEvents[Index].EventType = E_EventType.Trigger THEN
        FTriggerCount := FTriggerCount + 1;
    END_IF;
END_FOR;
FStepExecuted := TRUE;
END_METHOD

END_FUNCTION_BLOCK

// ---- SelfTests/TestCases/TestSuite_RunControlLifecycle/Test_RunControlNormalLifecycle.TcPOU
{region 'Documentation'}
(*!
<summary>Runs the real root twice, checking Suite aggregation and fresh finalization after lifecycle Reset.</summary>
<description>

Independent observations

Each script step calls the subject once. The helper sees the previous child snapshots,
then ProcessTestSuites applies the new ones; counters must reflect them in that same call.
Completion requires both children and the helper. Passed/Failed is finalized in Completing.

Repeated lifecycle

Initialize is called only for the first run. The second run uses RequestReset and RequestStart
with the original collection and service bindings. FirstChildResult selects Passed or Failed
for the first run; the second run is always Passed to expose retained result/finalization data.
CompletionDelay is zero here; duration and clock-failure qualification belong to separate tests.

Event evidence

One local capture retains both runs. The test checks one Result and Aggregation per run,
their structured context and compact JSON counts/runtime, and the later Completed anchor.
Expected payloads are built from scenario values, not the production event factory.
</description>
*)
{endregion}
FUNCTION_BLOCK Test_RunControlNormalLifecycle EXTENDS TestCaseBase
VAR_INPUT
    FirstChildResult : E_Result := E_Result.Passed; //! Passed or Failed for the first run; held constant by the containing test Suite.
END_VAR
VAR
    FSubject : RunControlLifecycleProbe;
    FHelper : SuiteOrchestratorDouble;
    FControl : ST_RunControl;
    FCapture : EventBuffer;
    FEvents : ARRAY[1..CaptureLength] OF ST_Event;
    FCaptureFifo : ST_FifoStatus;
    FCaptureStatus : ST_EventBufferStatus;
    FStep : INT;
    FRun : INT := 1;
    FRunChildResult : E_Result;
    FRunRuntime : ARRAY[1..RunCount] OF TIME;
    FStepChecked : BOOL;
    FStatePath : AssertTrue;
    FStatePathMatches : BOOL := TRUE;
    FTaskMapping : AssertTrue;
    FTaskMappingMatches : BOOL := TRUE;
    FOwnerResult : AssertTrue;
    FOwnerResultMatches : BOOL := TRUE;
    FStatusCounters : AssertTrue;
    FStatusCountersMatches : BOOL := TRUE;
    FCallOrder : AssertTrue;
    FCallOrderMatches : BOOL := TRUE;
    FReadiness : AssertTrue;
    FReadinessMatches : BOOL := TRUE;
    FFinalEvents : AssertTrue;
    FFinalEventsMatches : BOOL := TRUE;
    FAggregationPayload : AssertTrue;
    FAggregationPayloadMatches : BOOL := TRUE;
    FCaptureIntegrity : AssertTrue;
    FCaptureIntegrityMatches : BOOL := TRUE;
END_VAR
VAR CONSTANT
    CaptureLength : UINT := 64;
    ExpectedChildCount : UINT := 2;
    RunCount : INT := 2;
    Setup : INT := 0;
    ChildrenReady : INT := 1;
    ResetFinished : INT := 2;
    StartReady : INT := 3;
    StartRequested : INT := 4;
    FirstChildCompleted : INT := 5;
    AllChildrenCompleted : INT := 6;
    WaitForHelper : INT := 7;
    OwnerCompleting : INT := 8;
    OwnerCompleted : INT := 9;
    HoldCompleted : INT := 10;
    StartWithoutReset : INT := 11;
    StepsPerRun : INT := 12;
END_VAR

SUPER^();

{region 'Documentation'}
(*!
<summary>Contributes only the checking Assertions, not the intentionally controlled subject results.</summary>
*)
{endregion}
METHOD PROTECTED AggregateResults
VAR_INPUT
    Aggregator : I_ResultAggregator; //! Borrowed result sink owned by the outer Test Case; add this test's checking Assertions without resetting or retaining the sink.
END_VAR
Aggregator.AddProvider(Provider := FStatePath);
Aggregator.AddProvider(Provider := FTaskMapping);
Aggregator.AddProvider(Provider := FOwnerResult);
Aggregator.AddProvider(Provider := FStatusCounters);
Aggregator.AddProvider(Provider := FCallOrder);
Aggregator.AddProvider(Provider := FReadiness);
Aggregator.AddProvider(Provider := FFinalEvents);
Aggregator.AddProvider(Provider := FAggregationPayload);
Aggregator.AddProvider(Provider := FCaptureIntegrity);
END_METHOD

{region 'Documentation'}
(*!
<summary>Checks both retained run logs against independently constructed final payload and ordering expectations.</summary>
*)
{endregion}
METHOD PRIVATE CheckFinalEvents
VAR
    Index : UINT;
    ResultCount : INT;
    AggregationCount : INT;
    CompletedCount : INT;
    ExpectedFinalCount : INT;
    ExpectedCompletedCount : INT;
    ExpectedResult : E_Result;
    ExpectedMessage : STRING(GVL_Constants.MessageLength);
    ResultSequence : UDINT;
    AggregationSequence : UDINT;
END_VAR
FFinalEventsMatches := TRUE;
FAggregationPayloadMatches := TRUE;
ExpectedFinalCount := FRun - 1 + BOOL_TO_INT(FStep >= OwnerCompleting);
ExpectedCompletedCount := FRun - 1 + BOOL_TO_INT(FStep >= OwnerCompleted);
FOR Index := 1 TO FCaptureFifo.ElementCount DO
    FFinalEventsMatches := FFinalEventsMatches
        AND (FEvents[Index].OwnerScope = E_OwnerScope.RunControl)
        AND (FEvents[Index].Name = 'LifecycleSubject');
    CASE FEvents[Index].EventType OF
        E_EventType.Result:
            ResultCount := ResultCount + 1;
            ExpectedResult := E_Result.Passed;
            IF ResultCount = 1 THEN
                ExpectedResult := FirstChildResult;
            END_IF;
            FFinalEventsMatches := FFinalEventsMatches
                AND (FEvents[Index].Result = ExpectedResult)
                AND (FEvents[Index].State = E_State.Completing)
                AND (FEvents[Index].ResourceName = 'Fixture')
                AND (FEvents[Index].Severity = E_EventSeverity.Info)
                AND (CompletedCount = ResultCount - 1)
                AND (AggregationCount = ResultCount - 1);
            ResultSequence := FEvents[Index].SequenceId;
        E_EventType.Aggregation:
            AggregationCount := AggregationCount + 1;
            IF AggregationCount > RunCount THEN
                FAggregationPayloadMatches := FALSE;
                CONTINUE;
            END_IF;
            ExpectedResult := E_Result.Passed;
            IF AggregationCount = 1 THEN
                ExpectedResult := FirstChildResult;
            END_IF;
            IF ExpectedResult = E_Result.Failed THEN
                ExpectedMessage := '{"total":2,"inactive":0,"idle":0,"running":0,"completed":2,"passed":1,"failed":1,"error":0,"runtime":';
            ELSE
                ExpectedMessage := '{"total":2,"inactive":0,"idle":0,"running":0,"completed":2,"passed":2,"failed":0,"error":0,"runtime":';
            END_IF;
            ExpectedMessage := CONCAT(ExpectedMessage, UDINT_TO_STRING(TIME_TO_UDINT(FRunRuntime[AggregationCount])));
            ExpectedMessage := CONCAT(ExpectedMessage, ',"lostEvents":0}');
            FAggregationPayloadMatches := FAggregationPayloadMatches
                AND (FEvents[Index].Message = ExpectedMessage)
                AND (FEvents[Index].Result = ExpectedResult)
                AND (FEvents[Index].State = E_State.Completing)
                AND (FEvents[Index].ResourceName = '')
                AND (FEvents[Index].Severity = E_EventSeverity.Info);
            AggregationSequence := FEvents[Index].SequenceId;
            FFinalEventsMatches := FFinalEventsMatches
                AND (ResultCount = AggregationCount)
                AND (ResultSequence < AggregationSequence)
                AND (CompletedCount = AggregationCount - 1);
        E_EventType.StateTransition:
            IF FEvents[Index].State = E_State.Completed THEN
                CompletedCount := CompletedCount + 1;
                FFinalEventsMatches := FFinalEventsMatches
                    AND (ResultCount = CompletedCount)
                    AND (AggregationCount = CompletedCount)
                    AND (AggregationSequence < FEvents[Index].SequenceId);
            END_IF;
    END_CASE;
END_FOR;
FFinalEventsMatches := FFinalEventsMatches
    AND (ResultCount = ExpectedFinalCount)
    AND (AggregationCount = ExpectedFinalCount)
    AND (CompletedCount = ExpectedCompletedCount);
END_METHOD

{region 'Documentation'}
(*!
<summary>Initializes the checking Assertions; the scenario explicitly initializes its isolated subject.</summary>
*)
{endregion}
METHOD PROTECTED Configure
FPreparationStateCount := 0;
FTestStateCount := RunCount * StepsPerRun;
FStatePath.Initialize(Parent := THIS^,
    AssertionName := 'StatePath');
FTaskMapping.Initialize(Parent := THIS^,
    AssertionName := 'TaskMapping');
FOwnerResult.Initialize(Parent := THIS^,
    AssertionName := 'OwnerResult');
FStatusCounters.Initialize(Parent := THIS^,
    AssertionName := 'StatusCounters');
FCallOrder.Initialize(Parent := THIS^,
    AssertionName := 'CallOrder');
FReadiness.Initialize(Parent := THIS^,
    AssertionName := 'Readiness');
FFinalEvents.Initialize(Parent := THIS^,
    AssertionName := 'FinalEvents');
FAggregationPayload.Initialize(Parent := THIS^,
    AssertionName := 'AggregationPayload');
FCaptureIntegrity.Initialize(Parent := THIS^,
    AssertionName := 'CaptureIntegrity');
END_METHOD

